  def clear_socket_buffer(gripper_socket="1", read_timeout = 0.1):
      rq_comm_clear_socket_buffer_enabled[rq_socket_to_index(gripper_socket)] = True
  end

  def rq_gripper_id_to_ascii(gripper_id):
      if(gripper_id == "1"):
          return 57
      elif(gripper_id == "2"):
          return 50
      elif(gripper_id == "3"):
          return 51
      elif(gripper_id == "4"):
          return 52
      end
  end

      def scale(value, rawRange, scaledRange):
          def computeSlope(inputRange, outputRange):
              outputRangeDelta = outputRange[1] - outputRange[0]
              inputRangeDelta = inputRange[1] - inputRange[0]

              if (inputRangeDelta == 0):
                  return 0
              else:
                  return outputRangeDelta / inputRangeDelta
              end
          end

          def computeIntercept(slope, inputRange, outputRange):
              return outputRange[0] - (slope * inputRange[0])
          end

          def clipScaledValue(outputScaledValue, outputRange):
              if (outputRange[0] < outputRange[1]):
                  return clipWhenLowerLimitIsLessThanHigher(outputScaledValue, outputRange)
              else:
                  return clipWhenLowerLimitIsGreaterThanHigherLimit(outputScaledValue, outputRange)
              end
          end

          def clipWhenLowerLimitIsGreaterThanHigherLimit(outputScaledValue, outputRange):
              if (outputScaledValue < outputRange[1]):
                  return outputRange[1]
              elif (outputScaledValue > outputRange[0]):
                  return outputRange[0]
              else:
                  return outputScaledValue
              end
          end

          def clipWhenLowerLimitIsLessThanHigher(outputScaledValue, outputRange):
              if (outputScaledValue < outputRange[0]):
                  return outputRange[0]
              elif (outputScaledValue > outputRange[1]):
                  return outputRange[1]
              else:
                  return outputScaledValue
              end
          end

          slope = computeSlope(rawRange, scaledRange)
          intercept = computeIntercept(slope, rawRange, scaledRange)
          scaledValue = slope * value + intercept
          return clipScaledValue(scaledValue, scaledRange)
      end

      def limit(value, range):
          return scale(value, range, range)
      end


  rq_init_comm_if_connected(9, "1")
  rq_init_comm_if_connected(2, "2")
  rq_init_comm_if_connected(3, "3")
  rq_init_comm_if_connected(4, "4")
  rq_print_connected_grippers()
  rq_gripper_communication_thread = run rq_gripper_communication()
  set_closed_norm(97.6470588235294, "1")
  set_open_norm(1.1764705882352942, "1")
  set_closed_mm(0.0, "1")
  set_open_mm(53.0, "1")
  set_closed_norm(100.0, "2")
  set_open_norm(0.0, "2")
  set_closed_mm(0.0, "2")
  set_open_mm(50.0, "2")
  set_closed_norm(100.0, "3")
  set_open_norm(0.0, "3")
  set_closed_mm(0.0, "3")
  set_open_mm(50.0, "3")
  set_closed_norm(100.0, "4")
  set_open_norm(0.0, "4")
  set_closed_mm(0.0, "4")
  set_open_mm(50.0, "4")
  rq_current_limit_enabled = False
  while(not rq_gripper_communication_thread_started):
      sleep(0.008)
  end
  # end: URCap Installation Node
  global AMR_Position=struct(position_identifier=0, x1=0, x2=0, y1=0, y2=0, theta1=0, theta2=0)
  global CAM_Pose=p[0,0,0,0,0,0]
  global CAM_Relation=""
  global CMD_Abort=  False
  global CMD_Clear=  False
  global CMD_Reset=  False
  global CMD_Start=  False
  global CMD_Suspend=  False
  global CMD_Unhold=  False
  global CMD_Unsuspend=  False
  global CNT_Rack_Output=0
  global FNC_Freedrive=  False
  global PRC_TubCounter=0
  global STP=0
  global easyPickCount_4=0
  global easyPickCount_7=0
  global easyPickNoObj_4=0
  global easyPickNoObj_7=0
  global easyPickParts_4=0
  global easyPickParts_7=0
  global TMR_Barcode=0
  global Container_mid_1_p=p[-.379239199143, -.127191311915, .299999999998, .000000000046, -.000000000021, -1.247199999994]
  global Container_mid_1_q=[-2.477408934449926, -1.2969853503591224, -1.875639182904262, -1.539621866126728, 1.5731943360401213, -2.8009955944022717]
  global trigger_otw_p=p[-.364831738276, -.163967193938, .343299997821, .000000000046, -.000000000020, -1.148401333327]
  global trigger_otw_q=[-2.378283213085033, -1.2994862387706814, -1.7634300687554951, -1.6493302004167063, 1.573123683454141, -2.8011223671816943]
  global Waypoint_54_p=p[.008800512419, -.547926542621, .402696567415, -.589884378425, -.007228654778, -.061268144704]
  global Waypoint_54_q=[-1.2044575850116175, -1.3416667741588135, -1.8272563219070435, -0.9884541195682068, 1.3621035814285278, -2.7712565104113978]
  global Waypoint_77_p=p[-.178371829612, -.433927395311, .368082383916, -.086593488055, .704679941724, -.007869906074]
  global Waypoint_77_q=[-1.265390698109762, -1.3355963987163086, -1.7944865226745605, -1.7402602634825648, 0.8780410885810852, -2.7713127771960657]
  global Waypoint_83_p=p[.008800512419, -.547926542621, .402696567415, -.589884378425, -.007228654778, -.061268144704]
  global Waypoint_83_q=[-1.2044575850116175, -1.3416667741588135, -1.8272563219070435, -0.9884541195682068, 1.3621035814285278, -2.7712565104113978]
  global Waypoint_84_p=p[-.178371829612, -.433927395311, .368082383916, -.086593488055, .704679941724, -.007869906074]
  global Waypoint_84_q=[-1.265390698109762, -1.3355963987163086, -1.7944865226745605, -1.7402602634825648, 0.8780410885810852, -2.7713127771960657]
  global Vial_above_1_p=p[.017105793010, -.652093028359, .184920586844, .000000000272, .000000000270, 1.564063451276]
  global Vial_above_1_q=[-1.3375440709712851, -1.9618096977868804, -1.4665759083780685, -1.2837941559171444, 1.5732503672317195, -4.47276330421513]
  global Vial_pick_poi_1_p=p[.017105792852, -.648922724010, .093307568731, .000000000271, .000000000270, 1.564063451276]
  global Vial_pick_poi_1_q=[-1.3366329456391917, -2.0375277831965413, -1.6071432798879028, -1.0675084332049813, 1.57309887265915, -4.471135348858068]
  global Waypoint_86_p=p[.019227646885, -.648669633640, .184920586950, .000000000000, .000000000000, .024063451426]
  global Waypoint_86_q=[-1.3331129109407733, -1.9540750545686123, -1.4775914902901128, -1.280581784992414, 1.5733500744865856, -2.928303704452631]
  global Waypoint_87_p=p[-.032361834699, -.348336136197, .391475576335, -.000008499254, .000014589902, -.004651426820]
  global Waypoint_87_q=[-1.2709335019096129, -1.1914598663441005, -1.708995335060501, -1.8117888533498316, 1.5729683532263925, -2.8379347397710237]
  global Vial_3FG_plac_1_p=p[-.031858676359, -.349402499566, .145301120695, .000000000000, .000000000000, .000000000000]
  global Vial_3FG_plac_1_q=[-1.2723975525801707, -1.252376585823825, -2.3128114007049496, -1.1470592278900167, 1.5730548099411423, -2.8414815174610535]
  global Waypoint_88_p=p[-.032361834699, -.348336136197, .391475576335, -.000008499254, .000014589902, -.004651426820]
  global Waypoint_88_q=[-1.2709335019096129, -1.1914598663441005, -1.708995335060501, -1.8117888533498316, 1.5729683532263925, -2.8379347397710237]
  global cap_dump_1_p=p[-.139168676487, -.420163541420, .146096395183, .000000000000, .000000000000, .000000000000]
  global cap_dump_1_q=[-1.584588644510994, -1.5093464179777323, -2.1118449369620347, -1.091059703602438, 1.5728943834877336, -3.154014906686923]
  global Waypoint_89_p=p[-.032361834699, -.348336136197, .391475576335, -.000008499254, .000014589902, -.004651426820]
  global Waypoint_89_q=[-1.2709335019096129, -1.1914598663441005, -1.708995335060501, -1.8117888533498316, 1.5729683532263925, -2.8379347397710237]
  global Vial_3FG_plac_2_p=p[-.031858676359, -.349402499566, .145301120695, .000000000000, .000000000000, .000000000000]
  global Vial_3FG_plac_2_q=[-1.2723975525801707, -1.252376585823825, -2.3128114007049496, -1.1470592278900167, 1.5730548099411423, -2.8414815174610535]
  global Waypoint_90_p=p[-.032361834699, -.348336136197, .391475576335, -.000008499254, .000014589902, -.004651426820]
  global Waypoint_90_q=[-1.2709335019096129, -1.1914598663441005, -1.708995335060501, -1.8117888533498316, 1.5729683532263925, -2.8379347397710237]
  global cap_dump_2_p=p[-.139168676487, -.420163541420, .146096395183, .000000000000, .000000000000, .000000000000]
  global cap_dump_2_q=[-1.584588644510994, -1.5093464179777323, -2.1118449369620347, -1.091059703602438, 1.5728943834877336, -3.154014906686923]
  global Waypoint_91_p=p[-.032361834699, -.348336136197, .391475576335, -.000008499254, .000014589902, -.004651426820]
  global Waypoint_91_q=[-1.2709335019096129, -1.1914598663441005, -1.708995335060501, -1.8117888533498316, 1.5729683532263925, -2.8379347397710237]
  global Vial_liq_abov_1_p=p[-.025303660977, -.338758622354, .426628485936, -1.315858642253, .800043520260, -.928295855026]
  global Vial_liq_abov_1_q=[-0.3789628187762659, -1.5149522957256814, -2.263045310974121, 0.7870649534412841, -0.750984017048971, -3.2237566153155726]
  global Vial_liq_pick_3_p=p[-.002660428945, -.335984893034, .159389832934, -1.150456778400, .673175527684, -1.010612657503]
  global Vial_liq_pick_3_q=[-0.3660772482501429, -1.4503649038127442, -2.4056053161621094, -1.994692941705221, 0.8039668202400208, -0.2508929411517542]
  global Vial_liq_pick_4_p=p[-.041402486291, -.356791603314, .125395323246, -1.143483969075, .651070210027, -.878721885453]
  global Vial_liq_pick_4_q=[-0.4426233705502476, -1.437252121513727, -2.551930962114307, -1.776528229806984, 0.6562026234073748, -0.43018811960029524]
  global Vial_liq_abov_2_p=p[-.025303660977, -.338758622354, .426628485936, -1.315858642253, .800043520260, -.928295855026]
  global Vial_liq_abov_2_q=[-0.3789628187762659, -1.5149522957256814, -2.263045310974121, 0.7870649534412841, -0.750984017048971, -3.2237566153155726]
  global Liquid_midway_1_p=p[.057575295009, -.583081747994, .306414980749, -1.351675548728, .120935756539, -.096908606303]
  global Liquid_midway_1_q=[-0.895174805318014, -1.7035466633238734, -2.380953073501587, 0.631549521083496, 0.7706599235534668, -2.9455552736865442]
  global shake_3_p=p[.057574880217, -.583085370269, .306422893466, -1.360996190983, -.155555042453, -.438136255921]
  global shake_3_q=[-0.8951800505267542, -1.7035466633238734, -2.380937099456787, 0.6315542894550782, 0.7706599235534669, -2.5394540616517496]
  global shake_4_p=p[.057581636113, -.583090570002, .306439684073, -1.308767904323, .368530312677, .214926493520]
  global shake_4_q=[-0.8951714674579065, -1.7035395107665003, -2.380906343460083, 0.6315504747578125, 0.7706480026245118, -3.3161255787892268]
  global drop_above_3_p=p[.268235025993, -.467784390499, .226219872376, -1.027832627524, -.430841408251, 1.004603115937]
  global drop_above_3_q=[-0.935645882283346, -1.6663371525206507, -2.4252893924713135, 0.41966931402172847, 1.8470635414123535, -3.4600217978106897]
  global drop_above_4_p=p[.219042229014, -.470775657081, .133754190740, -.313004595901, -.344395319364, 1.500564994056]
  global drop_above_4_q=[-1.0601594887284795, -1.70046459045642, -2.0799996233759863, -0.7243227230676759, 1.9429634314685202, -4.115129153870795]
  global liq_tran_3_p=p[.213067510942, -.469567035397, .100231043184, .251862243732, .217902579404, 1.592812335393]
  global liq_tran_3_q=[-0.7789645168037476, -1.822364827406652, -1.8643518410805573, -1.252158963840138, 1.3768134449520435, -3.9328333233290254]
  global drop_above_5_p=p[.219042229014, -.470775657081, .133754190740, -.313004595901, -.344395319364, 1.500564994056]
  global drop_above_5_q=[-1.0601594887284795, -1.70046459045642, -2.0799996233759863, -0.7243227230676759, 1.9429634314685202, -4.115129153870795]
  global Waypoint_92_p=p[.187119460405, -.493959476151, .133754190608, -.313004596540, -.344395317757, 1.500564993991]
  global Waypoint_92_q=[-1.1418328121400876, -1.7310553375189475, -2.033634768766424, -0.772026910513711, 1.958578934631971, -4.201588449364511]
  global liq_tran_4_p=p[.195957706507, -.493022614126, .100231042689, .160718757180, .109807038912, 1.525321508623]
  global liq_tran_4_q=[-0.881740380645474, -1.8244526267589851, -1.865100964490387, -1.1608866323693583, 1.4631433601076713, -3.973915130363038]
  global drop_above_6_p=p[.219042229014, -.470775657081, .133754190740, -.313004595901, -.344395319364, 1.500564994056]
  global drop_above_6_q=[-1.0601594887284795, -1.70046459045642, -2.0799996233759863, -0.7243227230676759, 1.9429634314685202, -4.115129153870795]
  global drop_above_7_p=p[.268235025993, -.467784390499, .226219872376, -1.027832627524, -.430841408251, 1.004603115937]
  global drop_above_7_q=[-0.935645882283346, -1.6663371525206507, -2.4252893924713135, 0.41966931402172847, 1.8470635414123535, -3.4600217978106897]
  global Liquid_midway_2_p=p[.057575295009, -.583081747994, .306414980749, -1.351675548728, .120935756539, -.096908606303]
  global Liquid_midway_2_q=[-0.895174805318014, -1.7035466633238734, -2.380953073501587, 0.631549521083496, 0.7706599235534668, -2.9455552736865442]
  global Vial_drop_abo_1_p=p[.000324902251, -.648569523142, .221894115667, -.873462921366, 1.165852672573, -1.482720593185]
  global Vial_drop_abo_1_q=[-1.0576906334721352, -2.393016994184633, -0.9236232851859159, -2.5729213042279273, 0.7903331288549689, -0.33286325848155585]
  global Vial_liq_drop_1_p=p[.001020867953, -.647659915585, .092915870838, -.834762611599, 1.081942994823, -1.540647900176]
  global Vial_liq_drop_1_q=[-1.0631954168193474, -2.4447642951220825, -1.128811017825127, -2.1983115491972294, 0.8130148661460634, -0.38984988696911316]
  global Vial_drop_abo_2_p=p[.000324902251, -.648569523142, .221894115667, -.873462921366, 1.165852672573, -1.482720593185]
  global Vial_drop_abo_2_q=[-1.0576906334721352, -2.393016994184633, -0.9236232851859159, -2.5729213042279273, 0.7903331288549689, -0.33286325848155585]
  global Spatula_otw_p=p[-.038472058237, -.263141484147, .425351216717, -.000441582511, -.000128175490, 3.034387645854]
  global Spatula_otw_q=[-1.1888947506684495, -1.0083288774886814, -1.7052227056065874, -1.9984805067363443, 1.5730180972985317, 0.48793409320312264]
  global pick_spat_L_abv_p=p[.239059466375, -.067212518441, .280720723617, .000017217488, -.000484427718, 3.106837214660]
  global pick_spat_L_abv_q=[0.292765616142962, -0.8565557553273315, -2.140199892763044, -1.715349495646084, 1.573623142106424, 1.8984976776985687]
  global spat_L_pick_p=p[.242468789885, -.067301915011, .193171208067, .000017217488, -.000484427718, 3.106837214657]
  global spat_L_pick_q=[0.2867414378807389, -0.8600077002089179, -2.3629148016312627, -1.4891831672860159, 1.5737695566221115, 1.8933890858591198]
  global spat_L_lift_p=p[.245402002494, -.067432373551, .289049296496, .000017217490, -.000484427724, 3.106837214657]
  global spat_L_lift_q=[0.2834351187564135, -0.8798320076811592, -2.1119436738532986, -1.7203314352121302, 1.573588313403067, 1.8891054681654005]
  global spat_L_side_p=p[.247133573905, -.017633681797, .289062935631, .000017217490, -.000484427724, 3.106837214657]
  global spat_L_side_q=[0.49719173575848863, -0.8582398211168538, -2.1182130454788215, -1.735610316654931, 1.5735817737572706, 2.1028402698705397]
  global spat_L_up_p=p[.247135508752, -.017665230822, .397130746165, .000017217490, -.000484427724, 3.106837214657]
  global spat_L_up_q=[0.49854946074076967, -0.9346239623559676, -1.808280269374471, -1.969158816463132, 1.5731020084036995, 2.1031742024348157]
  global spat_M_up_p=p[.244670000000, -.112000000000, .420343789747, .000026293990, -.000477463070, 3.067686800857]
  global spat_M_up_q=[0.09097498152209688, -1.0114245603211778, -1.718034632879454, -1.9826932847219538, 1.5730130135866505, 1.734554438783734]
  global spat_M_pick_p=p[.244673518506, -.111985070134, .192299022723, .000043885692, -.000001622442, 3.067686841404]
  global spat_M_pick_q=[0.08868170265231701, -0.9271392933223233, -2.343826449241451, -1.441236864368305, 1.5733923850045939, 1.7345552462242537]
  global spat_S_Up_7_p=p[.243228810603, -.161948321982, .423281604617, .000026293955, -.000477463064, 3.067686800854]
  global spat_S_Up_7_q=[-0.11182322368059516, -1.0716267311491734, -1.6854498186860427, -1.955120134033855, 1.5730106579635699, 1.5317349120701778]
  global spat_S_Pick_4_p=p[.245377020686, -.158668022535, .192285730279, .000026293985, -.000477463062, 3.067686800840]
  global spat_S_Pick_4_q=[-0.10087203759495189, -1.011188488703386, -2.311978084495874, -1.3890267520590838, 1.5735990551056096, 1.5450562970948172]
  global spat_S_Up_8_p=p[.252087445596, -.159242094834, .423281604617, .000026293954, -.000477463070, 3.067686800855]
  global spat_S_Up_8_q=[-0.09804692328730358, -1.0862987822056382, -1.6788706463996483, -1.9470242450550348, 1.5730147401359813, 1.5455107082823842]
  global spat_flatM_up_p=p[.241028517126, -.208127630016, .404671074680, .000026293951, -.000477463078, 3.067686800891]
  global spat_flatM_up_q=[-0.27878462628263456, -1.1217510366315881, -1.7121530048618725, -1.8783279876432832, 1.5731053960668042, 1.3649536117980254]
  global spat_flatM_pick_p=p[.241028983327, -.208057297586, .192270533170, .000026293950, -.000477463079, 3.067686800885]
  global spat_flatM_pick_q=[-0.2805687960562633, -1.1003763929487214, -2.271431297337675, -1.3404236887924883, 1.5734924238720627, 1.3653813047742556]
  global spat_flatS_up_p=p[.237651953780, -.253943828614, .403961222825, .000026293950, -.000477463092, 3.067686800841]
  global spat_flatS_up_q=[-0.42363550926974103, -1.1939944599502539, -1.6745915127240307, -1.843675057902054, 1.5731001874678698, 1.220082820532415]
  global spat_flatS_pick_p=p[.241325662334, -.251726327528, .192256842740, .000026293947, -.000477463087, 3.067686800841]
  global spat_flatS_pick_q=[-0.4144907797170738, -1.1967447109013012, -2.21926362252748, -1.2962499335425761, 1.5733885098427622, 1.2314402238866728]
  global spat_S_pick_p=p[.241585614619, -.158882677087, .191636172448, .000019478956, -.000483249177, 3.097147973434]
  global spat_S_pick_q=[-0.10320942227973173, -1.0007485193115802, -2.317947069452162, -1.3934956127505886, 1.5736112980229278, 1.5132597021160705]
  global spat_S_up_p=p[.248189103503, -.159371150053, .417088864416, .000026293966, -.000477463070, 3.067686800840]
  global spat_S_up_q=[-0.10007737460061872, -1.0730270029702904, -1.7018049146034766, -1.9373622285571734, 1.573045444550866, 1.5435422173047084]
  global Waypoint_7_p=p[-.472820924474, .292439826233, .207418370237, -.137787250486, 2.177332259632, -2.152029714756]
  global Waypoint_7_q=[-2.911134078210732, -1.90240864358569, -1.968768330510411, -2.500365101593811, 0.11427687110891149, 0.0958980389250167]
  global Waypoint_8_p=p[-.357612884176, -.251084817998, .212379799667, -.858181193174, 1.714832512191, -1.687547565568]
  global Waypoint_8_q=[-1.620834863369681, -1.8936194567376496, -1.9821394403832038, -2.4599791457905273, 0.6296693672615152, 0.07625365420707819]
  global Decapp_above_3_p=p[-.013480295948, -.359153355979, .266194408367, -.879653555922, 1.646336924805, -1.709111068605]
  global Decapp_above_3_q=[-0.9632157249872035, -2.0163405763031657, -1.5968194594157152, -2.6579215719847085, 1.251243398585566, 0.047906446502667066]
  global Decapp_place_3_p=p[-.013480295890, -.359153356055, .160907502384, -.879653554902, 1.646336919740, -1.709111066456]
  global Decapp_place_3_q=[-0.9633402410919709, -2.1541179572356635, -1.6937729380888573, -2.4232786481058053, 1.2517342187662468, 0.04818402956922263]
  global Decapp_above_4_p=p[-.013480295948, -.359153355979, .266194408367, -.879653555922, 1.646336924805, -1.709111068605]
  global Decapp_above_4_q=[-0.9632157249872035, -2.0163405763031657, -1.5968194594157152, -2.6579215719847085, 1.251243398585566, 0.047906446502667066]
  global Waypoint_78_p=p[-.051450028091, -.519555688329, .365718563414, -1.287302938145, 1.077637394477, -1.218524965834]
  global Waypoint_78_q=[-0.9214276262416012, -1.8899696965062578, -1.4939326452510562, -2.840015661555725, 0.5585157189668353, 0.033997638875617575]
  global Waypoint_10_p=p[-.466751210260, .252836712095, .259921246286, 1.042686976164, .439333316918, -1.691967798809]
  global Waypoint_10_q=[-3.022216346250036, -1.8383597675135919, -1.566977059184386, -2.046864464116096, 0.8487467526238, -2.4392912369481916]
  global Waypoint_9_p=p[-.538777454962, .370695704977, .175030018143, -.317104215445, 2.082346543003, -2.037631421082]
  global Waypoint_9_q=[-3.1158871966457857, -1.998548595120492, -1.941797010061462, -2.2703530575838844, -0.27573365931009164, -0.06926782177267654]
  global Powder_wayp1_p=p[-.472820924474, .292439826233, .207418370237, -.137787250486, 2.177332259632, -2.152029714756]
  global Powder_wayp1_q=[-2.911134078210732, -1.90240864358569, -1.968768330510411, -2.500365101593811, 0.11427687110891149, 0.0958980389250167]
  global Waypoint_2_p=p[-.357612884176, -.251084817998, .212379799667, -.858181193174, 1.714832512191, -1.687547565568]
  global Waypoint_2_q=[-1.620834863369681, -1.8936194567376496, -1.9821394403832038, -2.4599791457905273, 0.6296693672615152, 0.07625365420707819]
  global Postions_otw_p=p[-.010896578244, -.533368729951, .288851175116, -1.233738470894, 1.195331112012, -1.207314088469]
  global Postions_otw_q=[-0.898791023514228, -2.078490033037677, -1.4499891355755317, -2.7624416226992476, 0.6570218891920963, 0.02136606178275929]
  global cont_A_otw_p=p[.070238108556, -.655257851554, .184611566008, -1.090601381517, 1.404822685081, -1.413645380264]
  global cont_A_otw_q=[-0.990969136335913, -2.7123780097559784, -0.5772671651193146, -3.0005537851220403, 0.84719335943793, 0.020652463706785973]
  global cont_B_otw_p=p[.255895686750, -.501120003087, .157855243207, -1.209177187561, 1.209243088037, -1.209202949417]
  global cont_B_otw_q=[-0.5819602570351563, -2.5181180937953833, -1.0264696604583161, -2.7360726814058687, 0.9880932038785559, -0.004134033524621827]
  global cont_B_safe_p=p[.242897168204, -.501733713795, .237745474779, -1.209212324107, 1.209144328638, -1.209309913894]
  global cont_B_safe_q=[-0.5929699566143585, -2.4210115429142114, -0.9949203644592259, -2.8646436479104267, 0.976678899749076, -0.004020526358775811]
  global cont_C_otw_p=p[.319495487998, -.362719410364, .163846736977, -1.233784872294, 1.195277203291, -1.207325031551]
  global cont_C_otw_q=[-0.3611889651645974, -2.404603865546651, -1.2341573845076566, -2.650535279811077, 1.1944844573128257, 0.01638086594640864]
  global Waypoint_1_p=p[-.352029261722, -.424157832422, .472326578019, -.000004407962, .000020663369, -1.529709227737]
  global Waypoint_1_q=[-2.017015745614491, -1.7423968528991196, -1.0053357238485425, -1.9644715035904907, 1.5727249689896, -2.060727852912713]
  global Waypoint_5_p=p[.219993437017, -.447144142811, .462350040687, .000006087494, .000031090075, .000022232405]
  global Waypoint_5_q=[-0.8406239476037944, -1.5982534362206806, -1.1934200873248484, -1.9205794898315975, 1.5727336676986443, -2.4135960466995314]
  global place_2_home_p=p[-.352029261717, -.424157832411, .329197314759, -.000004407962, .000020663369, -1.529709227737]
  global place_2_home_q=[-2.017880982348384, -1.6708952803108668, -1.462293789471877, -1.5790150659586653, 1.5732060241635952, -2.059940179665328]
  global Waypoint_12_p=p[-.812560029877, -.415067232840, .258518340146, -1.257569567036, 1.159670338548, -1.145019586130]
  global Waypoint_12_q=[-2.3224548809497123, -2.3211405271930765, -1.1304722687551445, -2.8155296475017018, -0.8321758827962036, -0.007205995478960503]
  global Waypoint_18_p=p[-.813643087636, -.416224939441, .099970000000, -1.257570310935, 1.159676546330, -1.145010619029]
  global Waypoint_18_q=[-2.322494764677227, -2.501268559301314, -1.239250885783676, -2.5265468980680197, -0.831327849164623, -0.00732105677136996]
  global Waypoint_19_p=p[-.812560029269, -.415067232191, .079455005744, -1.257569567033, 1.159670338546, -1.145019586137]
  global Waypoint_19_q=[-2.3224951834453367, -2.5274729453886575, -1.2489176533831348, -2.4906644180980346, -0.8312252662037514, -0.007338111970053518]
  global TMR_Barcode_is_counting=False
  thread Timer_Thread():
    while (True):
      if (TMR_Barcode_is_counting):
        TMR_Barcode = TMR_Barcode + get_steptime()
      end
      sync()
    end
  end
  run Timer_Thread()
  def Sub_Vision_V18():
    $ 887 "Sub_Vision_V18" "noBreak"
    $ 888 "PreSettings"
    $ 889 "CAM_LM_Detected≔ False "
    global CAM_LM_Detected=  False
    $ 890 "CAM_Captures≔0"
    global CAM_Captures=0
    $ 891 "CAM_Pose≔p[0,0,0,0,0,0]"
    global CAM_Pose=p[0,0,0,0,0,0]
    $ 892 "CAM_LM_Refinmnt≔ False "
    global CAM_LM_Refinmnt=  False
    $ 893 "CAM_LM_Refined≔ False "
    global CAM_LM_Refined=  False
    $ 894 "CAM_LM_Deviatn≔p[0,0,0,0,0,0]"
    global CAM_LM_Deviatn=p[0,0,0,0,0,0]
    $ 895 "CAM_LM_ID≔0"
    global CAM_LM_ID=0
    $ 896 "CAM_Done≔ False "
    global CAM_Done=  False
    $ 897 "CAM_CNT_Obj≔0"
    global CAM_CNT_Obj=0
    $ 898 "CAM_Result = []"
    CAM_Result = []
    $ 899 "OBJ_Detected≔ False "
    global OBJ_Detected=  False
    $ 900 "FRM_Reference≔p[0,0,0,0,0,0]"
    global FRM_Reference=p[0,0,0,0,0,0]
    $ 901 "'=========='"
    # '=========='
    $ 902 "Switch Action"
    switch_1 = Action
    $ 903 "Case 13"
    if (13 == switch_1):
    elif (15 == switch_1):
      $ 1021 "Case 15"
    elif (131 == switch_1):
      $ 1067 "Case 131"
      $ 1068 "Read (SensoPart)"
      $ 1069 "Action_Info≔'search for landmark'"
      global Action_Info="search for landmark"
      $ 1070 "CAM_LM≔CAM_LMs[4]"
      global CAM_LM=CAM_LMs[4]
      $ 1071 "CAM_Relation≔CAM_LM.capture_relation"
      global CAM_Relation=CAM_LM.capture_relation
      $ 1072 "go to capture pose"
      $ 1075 "If ITM_ID≟1 and JIG≟7"
      if (ITM_ID == 1  and  JIG == 7):
        $ 1076 "PSE_T≔uLM_Cap_SSRack"
        global PSE_T=uLM_Cap_SSRack
      else:
        $ 1077 "ElseIf ITM_ID≟5 and JIG≟7"
        if (ITM_ID == 5  and  JIG == 7):
          $ 1078 "PSE_T≔FRM_Cap_SSRack"
          global PSE_T=FRM_Cap_SSRack
        else:
          $ 1081 "ElseIf ITM_ID≟1 and JIG≟15"
          if (ITM_ID == 1 and JIG == 15):
            $ 1082 "MoveJ"
            $ 1083 "Container_mid_1" "breakAfter"
            movej(get_inverse_kin(Container_mid_1_p, qnear=Container_mid_1_q), a=1.3962634015954636, v=1.0471975511965976, r=0.05)
            $ 1085 "PSE_T≔FRM_Container_const"
            global PSE_T=p[-0.5003348223692186,0.35061804815168285,0.41579001388808423,-5.092943187272062E-5,1.0145185065363121E-4,-2.764319258713288]
          else:
            $ 1086 "ElseIf ITM_ID≟1 and JIG≟21"
            if (ITM_ID == 1 and JIG == 21):
              $ 1088 "PSE_T≔FRM_PoTS_const"
              global PSE_T=p[-0.5403054403210852,-0.10910773999775857,0.4828,3.058497512721046E-6,2.3454853329357316E-5,-2.208510541952706]
            else:
              $ 1089 "ElseIf ITM_ID≟1 and JIG≟17"
              if (ITM_ID == 1 and JIG == 17):
                $ 1090 "MoveJ"
                $ 1091 "zero_scale()"
                zero_scale()
                $ 1092 "trigger_otw" "breakAfter"
                movej(get_inverse_kin(trigger_otw_p, qnear=trigger_otw_q), a=1.3962634015954636, v=1.0471975511965976, r=0.05)
                $ 1096 "PSE_T≔FRM_weigh_scale_const"
                global PSE_T=p[-0.3804866881697204,0.025744252835212,0.4723487455232425,-1.0445769542396123E-4,-1.924788411074358E-5,-2.1691978730572363]
              end
            end
          end
        end
      end
      $ 1097 "do_transition(PSE_T, keep_rxry=False)"
      do_transition(PSE_T, keep_rxry=False)
      $ 1098 "Set"
      set_tcp(p[0.0,0.0,0.161,3.1415,0.0,0.0])
      $ 1099 "MoveJ"
      $ 1100 "PSE_T" "breakAfter"
      movej(PSE_T, a=1.3962634015954636, v=1.7453292519943295)
      $ 1101 "CAM_Pose≔get_actual_tcp_pose()"
      global CAM_Pose= get_actual_tcp_pose ()
      $ 1102 "Loop  not CAM_Done and  not ERROR.FLAG and  not CMD_Stop"
      while (  not  CAM_Done  and    not  ERROR.FLAG  and    not  CMD_Stop):
        $ 1103 "adjust capture pose"
        $ 1104 "If CAM_LM_Detected and CAM_LM_Refinmnt"
        if (CAM_LM_Detected  and  CAM_LM_Refinmnt):
          $ 1105 "PSE_T≔p[0,0,0.300,0,0,0]"
          global PSE_T=p[0,0,0.300,0,0,0]
          $ 1106 "CAM_Pose≔PSE_T"
          global CAM_Pose=PSE_T
          $ 1107 "If  not is_reachable(FRM_Reference,[PSE_T])"
          if (  not  is_reachable(FRM_Reference,[PSE_T])):
            $ 1108 "Error"
            $ 1109 "set_error(ERROR_POSE_NOT_REACHABLE)"
            set_error(ERROR_POSE_NOT_REACHABLE)
          end
          $ 1110 "If  not ERROR.FLAG"
          if (  not  ERROR.FLAG):
            $ 1111 "MoveJ"
            $ 1112 "PSE_T" "breakAfter"
            set_tcp(p[0.0,0.0,0.161,0.0,0.0,0.0])
            movej(pose_trans(FRM_Reference, PSE_T), a=0.8726646259971648, v=1.3962634015954636)
            $ 1113 "CAM_LM_Refined≔ True "
            global CAM_LM_Refined=  True
          end
        else:
          $ 1114 "ElseIf  not CAM_LM_Detected and CAM_Captures>0"
          if (  not  CAM_LM_Detected  and  CAM_Captures>0):
            $ 1115 "MoveL"
            $ 1116 "If FRM_Reference≟p[0,0,0,0,0,0]"
            if (FRM_Reference == p[0,0,0,0,0,0]):
              $ 1117 "PSE_T≔get_random_pose(pose_ref=CAM_Pose, mode='cubic', range_max=[0.150,0.150,0.015])"
              global PSE_T=get_random_pose(pose_ref=CAM_Pose, mode="cubic", range_max=[0.150,0.150,0.015])
            else:
              $ 1122 "Else" "noBreak"
              $ 1123 "PSE_T≔get_random_pose(pose_ref=CAM_Pose, mode='rotation', range_max=[10,10,0])"
              global PSE_T=get_random_pose(pose_ref=CAM_Pose, mode="rotation", range_max=[10,10,0])
              $ 1124 "CAM_LM_Refined≔ True "
              global CAM_LM_Refined=  True
            end
            $ 1125 "If get_inverse_kin_has_solution(pose_trans(FRM_Reference, PSE_T))"
            if (get_inverse_kin_has_solution( pose_trans (FRM_Reference, PSE_T))):
              $ 1126 "Comment"
              # Comment
              $ 1127 "PSE_T" "breakAfter"
              set_tcp(p[0.0,0.0,0.161,3.1415,0.0,0.0])
              movel(pose_trans(FRM_Reference, PSE_T), a=0.03, v=0.05)
            else:
              $ 1128 "Else" "noBreak"
              $ 1129 "'If random pose is out of reach, set the initial cam pose'"
              # 'If random pose is out of reach, set the initial cam pose'
              $ 1130 "PSE_T≔CAM_Pose"
              global PSE_T=CAM_Pose
            end
          end
        end
        $ 1131 "Wait: 2.0"
        sleep(2.0)
        $ 1132 "trigger"
        $ 1133 "If ITM_ID≟1 and JIG≟7"
        if (ITM_ID == 1  and  JIG == 7):
          # begin: URCap Program Node
          #   Source: SensoPart VISOR Robotic, 2.0.6, SensoPart Industriesensorik GmbH
          #   Type: VISOR Trigger
          $ 1134 "# 1 VISOR Trigger"
          visor_changeJob(1, "Landmark_INVITE_2", 6000)
          visor_trigger(1, 6000, "arm")
          # end: URCap Program Node
        else:
          $ 1135 "ElseIf ITM_ID≟5 and JIG≟7"
          if (ITM_ID == 5  and  JIG == 7):
            # begin: URCap Program Node
            #   Source: SensoPart VISOR Robotic, 2.0.6, SensoPart Industriesensorik GmbH
            #   Type: VISOR Trigger
            $ 1136 "# 1 VISOR Trigger"
            visor_changeJob(1, "Landmark_INVITE_2", 6000)
            visor_trigger(1, 6000, "arm")
            # end: URCap Program Node
          else:
            $ 1137 "ElseIf ITM_ID≟13 and JIG≟7"
            if (ITM_ID == 13  and  JIG == 7):
              # begin: URCap Program Node
              #   Source: SensoPart VISOR Robotic, 2.0.6, SensoPart Industriesensorik GmbH
              #   Type: VISOR Trigger
              $ 1138 "# 1 VISOR Trigger"
              visor_changeJob(1, "Landmark_INVITE_2", 6000)
              visor_trigger(1, 6000, "arm")
              # end: URCap Program Node
            else:
              $ 1139 "ElseIf ITM_ID≟1 and JIG≟15"
              if (ITM_ID == 1 and JIG == 15):
                # begin: URCap Program Node
                #   Source: SensoPart VISOR Robotic, 2.0.6, SensoPart Industriesensorik GmbH
                #   Type: VISOR Trigger
                $ 1140 "# 1 VISOR Trigger"
                visor_changeJob(1, "Aztec_no_dot_pick", 6000)
                visor_trigger(1, 6000, "arm")
                # end: URCap Program Node
              else:
                $ 1141 "ElseIf ITM_ID≟1 and JIG≟21"
                if (ITM_ID == 1 and JIG == 21):
                  # begin: URCap Program Node
                  #   Source: SensoPart VISOR Robotic, 2.0.6, SensoPart Industriesensorik GmbH
                  #   Type: VISOR Trigger
                  $ 1142 "# 1 VISOR Trigger"
                  visor_changeJob(1, "PoTS", 6000)
                  visor_trigger(1, 6000, "arm")
                  # end: URCap Program Node
                else:
                  $ 1143 "ElseIf ITM_ID≟1 and JIG≟17"
                  if (ITM_ID == 1 and JIG == 17):
                    # begin: URCap Program Node
                    #   Source: SensoPart VISOR Robotic, 2.0.6, SensoPart Industriesensorik GmbH
                    #   Type: VISOR Trigger
                    $ 1144 "# 1 VISOR Trigger"
                    visor_changeJob(1, "Weigh_target", 6000)
                    visor_trigger(1, 6000, "arm")
                    # end: URCap Program Node
                  end
                end
              end
            end
          end
        end
        $ 1148 "TM_3D_Found≔visor_partsFound(1)"
        global TM_3D_Found= visor_partsFound (1)
        $ 1150 "If TM_3D_Found>0"
        if (TM_3D_Found>0):
          $ 1151 "CAM_LM_Detected≔ True "
          global CAM_LM_Detected=  True
          $ 1152 "CAM_Captures≔0"
          global CAM_Captures=0
        else:
          $ 1153 "Else" "noBreak"
          $ 1154 "CAM_LM_Detected≔ False "
          global CAM_LM_Detected=  False
          $ 1155 "CAM_Captures≔CAM_Captures+1"
          global CAM_Captures=CAM_Captures+1
        end
        $ 1160 "result"
        $ 1161 "If CAM_LM_Detected"
        if (CAM_LM_Detected):
          $ 1162 "If (CAM_LM_Refinmnt and CAM_LM_Refined) or  not CAM_LM_Refinmnt"
          if ((CAM_LM_Refinmnt  and  CAM_LM_Refined)  or    not  CAM_LM_Refinmnt):
            $ 1220 "If ITM_ID≟1 and JIG≟7"
            if (ITM_ID == 1  and  JIG == 7):
              $ 1221 "CAM_LM_SSRack≔visor_getPose3d(1, 0)"
              global CAM_LM_SSRack= visor_getPose3d (1, 0)
            else:
              $ 1222 "ElseIf ITM_ID≟5 and JIG≟7"
              if (ITM_ID == 5  and  JIG == 7):
                $ 1223 "CAM_LM_SSRack≔visor_getPose3d(1, 0)"
                global CAM_LM_SSRack= visor_getPose3d (1, 0)
              else:
                $ 1226 "ElseIf ITM_ID≟1 and JIG≟15"
                if (ITM_ID == 1 and JIG == 15):
                  $ 1227 "CAM_LM_cont≔visor_getPose3d(1, 0)"
                  global CAM_LM_cont= visor_getPose3d (1, 0)
                  $ 1228 "Trigger≔get_actual_tcp_pose()"
                  global Trigger= get_actual_tcp_pose ()
                else:
                  $ 1229 "ElseIf ITM_ID≟1 and JIG≟21"
                  if (ITM_ID == 1 and JIG == 21):
                    $ 1230 "CAM_LM_cont≔visor_getPose3d(1, 0)"
                    global CAM_LM_cont= visor_getPose3d (1, 0)
                    $ 1231 "Trigger≔get_actual_tcp_pose()"
                    global Trigger= get_actual_tcp_pose ()
                  else:
                    $ 1232 "ElseIf ITM_ID≟1 and JIG≟17"
                    if (ITM_ID == 1 and JIG == 17):
                      $ 1233 "CAM_LM_cont≔visor_getPose3d(1, 0)"
                      global CAM_LM_cont= visor_getPose3d (1, 0)
                      $ 1234 "Trigger≔get_actual_tcp_pose()"
                      global Trigger= get_actual_tcp_pose ()
                    end
                  end
                end
              end
            end
            $ 1235 "CAM_Done≔ True "
            global CAM_Done=  True
          end
        else:
          $ 1236 "ElseIf  not CAM_LM_Detected and CAM_Captures<CAM_PRM_Retries"
          if (  not  CAM_LM_Detected  and  CAM_Captures<CAM_PRM_Retries):
            $ 1237 "CAM_LM_Refined≔ False "
            global CAM_LM_Refined=  False
          else:
            $ 1238 "ElseIf CAM_Captures≥CAM_PRM_Retries"
            if (CAM_Captures >= CAM_PRM_Retries):
              $ 1239 "CAM_Done≔ True "
              global CAM_Done=  True
              $ 1240 "Error"
              $ 1241 "set_error(ERROR_NO_LANDMARK)"
              set_error(ERROR_NO_LANDMARK)
            end
          end
        end
      end
    elif (151 == switch_1):
      $ 1242 "Case 151"
      $ 1243 "Detect (SensoPart)"
      $ 1244 "go to capture pose"
      $ 1245 "FRM_Reference≔FRM_Cap_SSRack"
      global FRM_Reference=FRM_Cap_SSRack
      $ 1246 "PSE_T≔p[0,0,-0.00,0,0,0]"
      global PSE_T=p[0,0,-0.00,0,0,0]
      $ 1247 "do_transition(pose_trans(FRM_Reference, PSE_T), keep_rxry=False)"
      do_transition( pose_trans (FRM_Reference, PSE_T), keep_rxry=False)
      $ 1248 "JNT_Q≔get_actual_joint_positions()"
      global JNT_Q= get_actual_joint_positions ()
      $ 1249 "JNT_Q≔[JNT_Q[0], JNT_Q[1], JNT_Q[2], JNT_Q[3], JNT_Q[4], 0]"
      global JNT_Q=[JNT_Q[0], JNT_Q[1], JNT_Q[2], JNT_Q[3], JNT_Q[4], 0]
      $ 1250 "Set"
      set_tcp(p[0.0,0.0,0.161,3.1415,0.0,0.0])
      $ 1251 "movej(get_inverse_kin(pose_trans(FRM_Reference, PSE_T), qnear=JNT_Q))"
      movej(get_inverse_kin( pose_trans (FRM_Reference, PSE_T), qnear=JNT_Q))
      $ 1252 "CAM_Pose≔pose_trans(pose_inv(FRM_Reference), get_actual_tcp_pose())"
      global CAM_Pose= pose_trans ( pose_inv (FRM_Reference),  get_actual_tcp_pose ())
      $ 1253 "Loop  not CAM_Done and  not ERROR.FLAG and  not CMD_Stop"
      while (  not  CAM_Done  and    not  ERROR.FLAG  and    not  CMD_Stop):
        $ 1254 "If  not OBJ_Detected and CAM_Captures>0"
        if (  not  OBJ_Detected  and  CAM_Captures>0):
          $ 1255 "MoveL"
          $ 1256 "If FRM_Reference≟p[0,0,0,0,0,0]"
          if (FRM_Reference == p[0,0,0,0,0,0]):
            $ 1258 "PSE_T≔get_random_pose(pose_ref=CAM_Pose, mode='rotation', range_max=[15,15,0])"
            global PSE_T=get_random_pose(pose_ref=CAM_Pose, mode="rotation", range_max=[15,15,0])
          else:
            $ 1259 "Else" "noBreak"
            $ 1260 "PSE_T≔get_random_pose(pose_ref=CAM_Pose, mode='rotation', range_max=[10,10,0])"
            global PSE_T=get_random_pose(pose_ref=CAM_Pose, mode="rotation", range_max=[10,10,0])
          end
          $ 1261 "If get_inverse_kin_has_solution(pose_trans(FRM_Reference, PSE_T))"
          if (get_inverse_kin_has_solution( pose_trans (FRM_Reference, PSE_T))):
            $ 1262 "PSE_T" "breakAfter"
            set_tcp(p[0.0,0.0,0.161,3.1415,0.0,0.0])
            movel(pose_trans(FRM_Reference, PSE_T), a=0.03, v=0.05)
          else:
            $ 1263 "Else" "noBreak"
            $ 1264 "'If random pose is out of reach, set the initial cam pose'"
            # 'If random pose is out of reach, set the initial cam pose'
            $ 1265 "PSE_T≔CAM_Pose"
            global PSE_T=CAM_Pose
            $ 1266 "PSE_T" "breakAfter"
            set_tcp(p[0.0,0.0,0.161,3.1415,0.0,0.0])
            movel(pose_trans(FRM_Reference, PSE_T), a=0.03, v=0.05)
          end
        end
        $ 1267 "Wait: 0.5"
        sleep(0.5)
        $ 1268 "Set"
        set_tcp(p[0.0,0.0,0.161,3.1415,0.0,0.0])
        # begin: URCap Program Node
        #   Source: SensoPart VISOR Robotic, 2.0.6, SensoPart Industriesensorik GmbH
        #   Type: VISOR Trigger
        $ 1269 "# 1 VISOR Trigger"
        visor_changeJob(1, "Object Detection Single", 6000)
        visor_trigger(1, 6000, "arm")
        # end: URCap Program Node
        $ 1270 "If visor_isResponseOk(1)"
        if ( visor_isResponseOk (1)):
          $ 1271 "CAM_CNT_Obj≔visor_partsFound(1)"
          global CAM_CNT_Obj= visor_partsFound (1)
          $ 1272 "CAM_OBJ_Pose≔visor_getPose3d(1, 0)"
          global CAM_OBJ_Pose= visor_getPose3d (1, 0)
          $ 1273 "If CAM_CNT_Obj>0"
          if (CAM_CNT_Obj>0):
            $ 1274 "CAM_OBJ_Color≔visor_getAdditionalData(1, 0)"
            global CAM_OBJ_Color= visor_getAdditionalData (1, 0)
            $ 1275 "CAM_DetectScore≔to_num(visor_getAdditionalData(1, 1))/1000"
            global CAM_DetectScore=to_num( visor_getAdditionalData (1, 1))/1000
            $ 1276 "OBJ_Detected≔ True "
            global OBJ_Detected=  True
          end
        else:
          $ 1277 "Else" "noBreak"
          $ 1278 "CAM_Captures≔CAM_Captures+1"
          global CAM_Captures=CAM_Captures+1
        end
        $ 1279 "If OBJ_Detected"
        if (OBJ_Detected):
          $ 1280 "Get object data"
          $ 1281 "PRC_CntDetect≔0"
          global PRC_CntDetect=0
          $ 1282 "Loop PRC_CntDetect<CAM_CNT_Obj"
          while (PRC_CntDetect<CAM_CNT_Obj):
            $ 1283 "get object and jig number"
            $ 1284 "If ITM_ID≟1 and JIG≟7"
            if (ITM_ID == 1  and  JIG == 7):
              $ 1285 "FRM_Reference≔FRM_Cap_SSRack"
              global FRM_Reference=FRM_Cap_SSRack
            else:
              $ 1286 "ElseIf ITM_ID≟5 and JIG≟7"
              if (ITM_ID == 5  and  JIG == 7):
                $ 1287 "FRM_Reference≔uLM_Cap_SSRack"
                global FRM_Reference=uLM_Cap_SSRack
              end
            end
            $ 1290 "PSE_T≔pose_trans(pose_inv(FRM_Reference), CAM_OBJ_Pose)"
            global PSE_T= pose_trans ( pose_inv (FRM_Reference), CAM_OBJ_Pose)
            $ 1291 "CAM_Result.append(get_pattern_counter(PSE_T, 'X', pattern=[10, 5], patternsize=[0.181, 0.081]))"
            CAM_Result.append(get_pattern_counter(PSE_T, "X", pattern=[10, 5], patternsize=[0.181, 0.081]))
            $ 1292 "PRC_CntDetect≔PRC_CntDetect+1"
            global PRC_CntDetect=PRC_CntDetect+1
          end
          $ 1293 "CAM_Done≔ True "
          global CAM_Done=  True
        else:
          $ 1294 "ElseIf CAM_Captures≥CAM_PRM_Retries"
          if (CAM_Captures >= CAM_PRM_Retries):
            $ 1295 "CAM_Done≔ True "
            global CAM_Done=  True
          else:
            $ 1296 "Else" "noBreak"
            $ 1297 "CAM_Captures≔CAM_Captures+1"
            global CAM_Captures=CAM_Captures+1
          end
        end
      end
    end
    $ 1298 "'=========='"
    # '=========='
    $ 1299 "PostSettings"
    $ 1300 "FRM_Reference≔p[0,0,0,0,0,0]"
    global FRM_Reference=p[0,0,0,0,0,0]
    $ 1301 "Set"
    set_tcp(p[0.0,0.0,0.161,3.1415,0.0,0.0])
    $ 1302 "CAM_Pose≔p[0,0,0,0,0,0]"
    global CAM_Pose=p[0,0,0,0,0,0]
    $ 1303 "Action≔0"
    global Action=0
    $ 1304 "Action_Info≔''"
    global Action_Info=""
  end
  def Sub_AMR_MiR_V3():
    $ 1305 "Sub_AMR_MiR_V3" "noBreak"
    $ 1306 "PreSettings"
    $ 1307 "AMR_TargetList≔[1,2,3,4,5,6,21,22,23,24,31,32,33,34,35,36,37,38,41]"
    global AMR_TargetList=[1,2,3,4,5,6,21,22,23,24,31,32,33,34,35,36,37,38,41]
    $ 1308 "AMR_Done≔ False "
    global AMR_Done=  False
    $ 1309 "AMR_PosActual≔T2O_Current_Pos"
    global AMR_PosActual=modbus_get_signal_status("T2O_Current_Pos")
    $ 1310 "AMR_Attemps≔T2O_Nav_Attemps"
    global AMR_Attemps=modbus_get_signal_status("T2O_Nav_Attemps")
    $ 1311 "AMR_Battery≔MiR_Battery_Lvl"
    global AMR_Battery=modbus_get_signal_status("MiR_Battery_Lvl")
    $ 1312 "AMR_Charging≔(T2O_Charging≟1)"
    global AMR_Charging=(modbus_get_signal_status("T2O_Charging") == 1)
    $ 1313 "AMR_Position≔struct(position_identifier=T2O_Current_Pos, x1=MiR_Position_X1, x2=MiR_Position_X2, y1=MiR_Position_Y1, y2=MiR_Position_Y2, theta1=MiR_Theta_1, theta2=MiR_Theta_2) "
    global AMR_Position=struct(position_identifier=modbus_get_signal_status("T2O_Current_Pos"), x1=modbus_get_signal_status("MiR_Position_X1"), x2=modbus_get_signal_status("MiR_Position_X2"), y1=modbus_get_signal_status("MiR_Position_Y1"), y2=modbus_get_signal_status("MiR_Position_Y2"), theta1=modbus_get_signal_status("MiR_Theta_1"), theta2=modbus_get_signal_status("MiR_Theta_2"))
    $ 1314 "If MiR_Mode≠7"
    if (modbus_get_signal_status("MiR_Mode") != 7):
      $ 1315 "Error"
      $ 1316 "set_error(ERROR_AMR_WRONG_MODE)"
      set_error(ERROR_AMR_WRONG_MODE)
      $ 1317 "AMR_Done≔ True "
      global AMR_Done=  True
    end
    $ 1318 "'=========='"
    # '=========='
    $ 1319 "Switch STATE"
    switch_1 = STATE
    $ 1320 "Case 1"
    if (1 == switch_1):
      $ 1321 "stopping"
      $ 1322 "If T2O_Done≟1 and O2T_Acknowledge≟0"
      if (modbus_get_signal_status("T2O_Done") == 1  and  modbus_get_signal_status("O2T_Acknowledge") == 0):
        $ 1323 "Set O2T_Acknowledge=1"
        modbus_set_output_register("O2T_Acknowledge", 1)
      end
      $ 1324 "Set MiR_CMD_Stop=On"
      modbus_set_output_signal("MiR_CMD_Stop", True)
      $ 1325 "AMR_Position.position_identifier = 0"
      AMR_Position.position_identifier = 0
      $ 1326 "AMR_Done≔ True "
      global AMR_Done=  True
    elif (2 == switch_1):
      $ 1327 "Case 2"
      $ 1328 "stopped"
      $ 1329 "If MiR_State≠3 and MiR_State≠5"
      if (modbus_get_signal_status("MiR_State") != 3  and  modbus_get_signal_status("MiR_State") != 5):
        $ 1330 "Set MiR_CMD_Stop=Off"
        modbus_set_output_signal("MiR_CMD_Stop", False)
      end
    elif (3 == switch_1):
      $ 1331 "Case 3"
      $ 1332 "resetting"
      $ 1333 "Set O2T_Mis_Main=Off"
      modbus_set_output_signal("O2T_Mis_Main", False)
      $ 1334 "Set O2T_Mis_Charge=Off"
      modbus_set_output_signal("O2T_Mis_Charge", False)
      $ 1335 "If MiR_Mis_Queue>0"
      if (modbus_get_signal_status("MiR_Mis_Queue")>0):
        $ 1336 "Set MiR_CMD_Clear_Q=On"
        modbus_set_output_signal("MiR_CMD_Clear_Q", True)
        $ 1337 "Wait MiR_Mis_Queue≟0"
        while (not(modbus_get_signal_status("MiR_Mis_Queue") == 0)):
          sync()
        end
        $ 1338 "Set MiR_CMD_Clear_Q=Off"
        modbus_set_output_signal("MiR_CMD_Clear_Q", False)
      end
      $ 1339 "If MiR_Error_ID≠0"
      if (modbus_get_signal_status("MiR_Error_ID") != 0):
        $ 1340 "Set MiR_CMD_Clear_E=On"
        modbus_set_output_signal("MiR_CMD_Clear_E", True)
        $ 1341 "Wait MiR_Error_ID≟0"
        while (not(modbus_get_signal_status("MiR_Error_ID") == 0)):
          sync()
        end
        $ 1342 "Set MiR_CMD_Clear_E=Off"
        modbus_set_output_signal("MiR_CMD_Clear_E", False)
      end
      $ 1343 "Set O2T_Action=0"
      modbus_set_output_register("O2T_Action", 0)
      $ 1344 "Set O2T_Acknowledge=0"
      modbus_set_output_register("O2T_Acknowledge", 0)
      $ 1345 "Set O2T_Target_Pos=0"
      modbus_set_output_register("O2T_Target_Pos", 0)
      $ 1346 "Set O2T_Footprint=0"
      modbus_set_output_register("O2T_Footprint", 0)
      $ 1347 "Set O2T_ProtectOff=0"
      modbus_set_output_register("O2T_ProtectOff", 0)
      $ 1348 "Set O2T_Dock=0"
      modbus_set_output_register("O2T_Dock", 0)
      $ 1349 "AMR_Attemps≔0"
      global AMR_Attemps=0
      $ 1350 "AMR_PosTarget≔0"
      global AMR_PosTarget=0
      $ 1351 "AMR_Step≔0"
      global AMR_Step=0
      $ 1352 "AMR_AtTarget≔ False "
      global AMR_AtTarget=  False
      $ 1353 "If MiR_State≟4 or MiR_State≟3 or MiR_State≟10"
      if (modbus_get_signal_status("MiR_State") == 4  or  modbus_get_signal_status("MiR_State") == 3  or  modbus_get_signal_status("MiR_State") == 10):
        $ 1354 "AMR_Done≔ True "
        global AMR_Done=  True
      end
    elif (5 == switch_1):
      $ 1355 "Case 5"
      $ 1356 "starting"
      $ 1357 "If MiR_State≟4"
      if (modbus_get_signal_status("MiR_State") == 4):
        $ 1358 "Set MiR_CMD_Start=On"
        modbus_set_output_signal("MiR_CMD_Start", True)
        $ 1359 "Wait MiR_State≠4"
        while (not(modbus_get_signal_status("MiR_State") != 4)):
          sync()
        end
        $ 1360 "Set MiR_CMD_Start=Off"
        modbus_set_output_signal("MiR_CMD_Start", False)
        $ 1361 "AMR_Done≔ True "
        global AMR_Done=  True
      else:
        $ 1362 "ElseIf MiR_State≟10"
        if (modbus_get_signal_status("MiR_State") == 10):
          $ 1363 "'MiR in protective stop. Wait'"
          # 'MiR in protective stop. Wait'
          $ 1364 "AMR_Done≔ True "
          global AMR_Done=  True
        else:
          $ 1365 "ElseIf MiR_State≟3"
          if (modbus_get_signal_status("MiR_State") == 3):
            $ 1366 "AMR_Done≔ True "
            global AMR_Done=  True
          end
        end
      end
    elif (6 == switch_1):
      $ 1367 "Case 6"
      $ 1368 "execute"
      $ 1369 "AMR_AtTarget≔(AMR_PosActual≟AMR_PosTarget)"
      global AMR_AtTarget=(AMR_PosActual == AMR_PosTarget)
      $ 1370 "Switch AMR_Step"
      switch_2 = AMR_Step
      $ 1371 "Case 0"
      if (0 == switch_2):
        $ 1372 "If  not AMR_AtTarget"
        if (  not  AMR_AtTarget):
          $ 1373 "AMR_Step≔1"
          global AMR_Step=1
        else:
          $ 1374 "Else" "noBreak"
          $ 1375 "AMR_Done≔ True "
          global AMR_Done=  True
        end
      elif (1 == switch_2):
        $ 1376 "Case 1"
        $ 1377 "general Settings"
        $ 1378 "Set O2T_Acknowledge=0"
        modbus_set_output_register("O2T_Acknowledge", 0)
        $ 1379 "check for error"
        $ 1380 "If OBJ_Picked and MiR_State≟10"
        if (OBJ_Picked  and  modbus_get_signal_status("MiR_State") == 10):
          $ 1381 "Error"
          $ 1382 "set_error(ERROR_ROBOT_ARM_NOT_IN_HOME_POSE)"
          set_error(ERROR_ROBOT_ARM_NOT_IN_HOME_POSE)
          $ 1383 "Action≔0"
          global Action=0
        else:
          $ 1384 "ElseIf  not found_in_list(AMR_PosTarget, AMR_TargetList)"
          if (  not  found_in_list(AMR_PosTarget, AMR_TargetList)):
            $ 1385 "Error"
            $ 1386 "set_error(ERROR_UNKNOWN_POSE)"
            set_error(ERROR_UNKNOWN_POSE)
            $ 1387 "Action≔0"
            global Action=0
          end
        end
        $ 1388 "If MiR_State≟3"
        if (modbus_get_signal_status("MiR_State") == 3):
          $ 1389 "Set MiR_CMD_Start=Off"
          modbus_set_output_signal("MiR_CMD_Start", False)
          $ 1390 "Switch Action"
          switch_3 = Action
          $ 1391 "Case 51"
          if (51 == switch_3):
            $ 1392 "Charge"
            $ 1393 "'trigger the charging mission'"
            # 'trigger the charging mission'
            $ 1394 "'target pos is predefined'"
            # 'target pos is predefined'
            $ 1395 "Set O2T_Footprint=0"
            modbus_set_output_register("O2T_Footprint", 0)
            $ 1396 "Set O2T_Action=1"
            modbus_set_output_register("O2T_Action", 1)
            $ 1397 "If MiR_Mis_Queue≟0"
            if (modbus_get_signal_status("MiR_Mis_Queue") == 0):
              $ 1398 "Set O2T_Mis_Charge=On"
              modbus_set_output_signal("O2T_Mis_Charge", True)
              $ 1399 "Wait MiR_Mis_Queue≥1"
              while (not(modbus_get_signal_status("MiR_Mis_Queue") >= 1)):
                sync()
              end
              $ 1400 "Set O2T_Mis_Charge=Off"
              modbus_set_output_signal("O2T_Mis_Charge", False)
            end
          elif (52 == switch_3):
            $ 1401 "Case 52"
            $ 1402 "Navigate"
            $ 1403 "'trigger the standard missoin'"
            # 'trigger the standard missoin'
            $ 1404 "Set O2T_Footprint=AMR_FootprintID"
            modbus_set_output_register("O2T_Footprint", AMR_FootprintID)
            $ 1405 "Set O2T_Target_Pos=AMR_PosTarget"
            modbus_set_output_register("O2T_Target_Pos", AMR_PosTarget)
            $ 1406 "Set O2T_Action=2"
            modbus_set_output_register("O2T_Action", 2)
            $ 1407 "If MiR_Mis_Queue≟0"
            if (modbus_get_signal_status("MiR_Mis_Queue") == 0):
              $ 1408 "Set O2T_Mis_Main=On"
              modbus_set_output_signal("O2T_Mis_Main", True)
              $ 1409 "Wait MiR_Mis_Queue≥1"
              while (not(modbus_get_signal_status("MiR_Mis_Queue") >= 1)):
                sync()
              end
              $ 1410 "Set O2T_Mis_Main=Off"
              modbus_set_output_signal("O2T_Mis_Main", False)
            end
          end
        else:
          $ 1411 "ElseIf MiR_State≟4"
          if (modbus_get_signal_status("MiR_State") == 4):
            $ 1412 "Set MiR_CMD_Start=On"
            modbus_set_output_signal("MiR_CMD_Start", True)
          else:
            $ 1413 "ElseIf MiR_State≟5"
            if (modbus_get_signal_status("MiR_State") == 5):
              $ 1414 "AMR_Step≔2"
              global AMR_Step=2
            else:
              $ 1415 "ElseIf MiR_State≟10"
              if (modbus_get_signal_status("MiR_State") == 10):
                $ 1416 "'AMR still in safeguard stop'"
                # 'AMR still in safeguard stop'
              end
            end
          end
        end
      elif (2 == switch_2):
        $ 1417 "Case 2"
        $ 1418 "acknowledge handshake"
        $ 1419 "If T2O_Done≟1 and O2T_Acknowledge≟0"
        if (modbus_get_signal_status("T2O_Done") == 1  and  modbus_get_signal_status("O2T_Acknowledge") == 0):
          $ 1420 "Set O2T_Acknowledge=1"
          modbus_set_output_register("O2T_Acknowledge", 1)
        else:
          $ 1421 "ElseIf T2O_Done≟0 and O2T_Acknowledge≟1"
          if (modbus_get_signal_status("T2O_Done") == 0  and  modbus_get_signal_status("O2T_Acknowledge") == 1):
            $ 1422 "Set O2T_Acknowledge=0"
            modbus_set_output_register("O2T_Acknowledge", 0)
            $ 1423 "AMR_AtTarget≔(AMR_PosActual≟AMR_PosTarget)"
            global AMR_AtTarget=(AMR_PosActual == AMR_PosTarget)
            $ 1424 "AMR_Done≔ True "
            global AMR_Done=  True
          end
        end
      end
      $ 1425 "translate errors"
      $ 1426 "If AMR_Done"
      if (AMR_Done):
        $ 1427 "Switch T2O_Error_ID"
        switch_2 = modbus_get_signal_status("T2O_Error_ID")
        $ 1428 "Case 2003"
        if (2003 == switch_2):
          $ 1429 "error"
          $ 1430 "set_error(ERROR_NOT_DOCKED)"
          set_error(ERROR_NOT_DOCKED)
        elif (2007 == switch_2):
          $ 1431 "Case 2007"
          $ 1432 "error"
          $ 1433 "set_error(ERROR_NOT_REACHABLE_TARGET)"
          set_error(ERROR_NOT_REACHABLE_TARGET)
        elif (2008 == switch_2):
          $ 1434 "Case 2008"
          $ 1435 "error"
          $ 1436 "set_error(ERROR_CHARGING_NOT_STARTED)"
          set_error(ERROR_CHARGING_NOT_STARTED)
        end
      end
    elif (7 == switch_1):
      $ 1437 "Case 7"
      $ 1438 "completing"
      $ 1439 "If MiR_Mis_Queue>0"
      if (modbus_get_signal_status("MiR_Mis_Queue")>0):
        $ 1440 "Set MiR_CMD_Abort=On"
        modbus_set_output_signal("MiR_CMD_Abort", True)
        $ 1441 "Wait MiR_Mis_Queue≟0"
        while (not(modbus_get_signal_status("MiR_Mis_Queue") == 0)):
          sync()
        end
        $ 1442 "Set MiR_CMD_Abort=Off"
        modbus_set_output_signal("MiR_CMD_Abort", False)
      end
      $ 1443 "If MiR_State≟3 or MiR_State≟10"
      if (modbus_get_signal_status("MiR_State") == 3  or  modbus_get_signal_status("MiR_State") == 10):
        $ 1444 "AMR_Done≔ True "
        global AMR_Done=  True
      end
    elif (9 == switch_1):
      $ 1445 "Case 9"
      $ 1446 "holding"
      $ 1447 "Set MiR_CMD_Abort=On"
      modbus_set_output_signal("MiR_CMD_Abort", True)
      $ 1448 "If MiR_State≟3 or MiR_State≟10"
      if (modbus_get_signal_status("MiR_State") == 3  or  modbus_get_signal_status("MiR_State") == 10):
        $ 1449 "Set MiR_CMD_Abort=Off"
        modbus_set_output_signal("MiR_CMD_Abort", False)
        $ 1450 "AMR_Done≔ True "
        global AMR_Done=  True
      end
    elif (11 == switch_1):
      $ 1451 "Case 11"
      $ 1452 "unholding"
      $ 1453 "Set MiR_CMD_Start=On"
      modbus_set_output_signal("MiR_CMD_Start", True)
      $ 1454 "If MiR_State≠4"
      if (modbus_get_signal_status("MiR_State") != 4):
        $ 1455 "Set MiR_CMD_Start=Off"
        modbus_set_output_signal("MiR_CMD_Start", False)
        $ 1456 "AMR_Step≔0"
        global AMR_Step=0
        $ 1457 "AMR_Done≔ True "
        global AMR_Done=  True
      end
    elif (12 == switch_1):
      $ 1458 "Case 12"
      $ 1459 "suspending"
      $ 1460 "'none'"
      # 'none'
    elif (14 == switch_1):
      $ 1461 "Case 14"
      $ 1462 "unsuspending"
      $ 1463 "'none'"
      # 'none'
    elif (15 == switch_1):
      $ 1464 "Case 15"
      $ 1465 "aborting"
      $ 1466 "Set MiR_CMD_Abort=On"
      modbus_set_output_signal("MiR_CMD_Abort", True)
      $ 1467 "Wait MiR_State≟3"
      while (not(modbus_get_signal_status("MiR_State") == 3)):
        sync()
      end
      $ 1468 "Set MiR_CMD_Abort=Off"
      modbus_set_output_signal("MiR_CMD_Abort", False)
    elif (17 == switch_1):
      $ 1469 "Case 17"
      $ 1470 "clearing"
      $ 1471 "If MiR_Error_ID≠0"
      if (modbus_get_signal_status("MiR_Error_ID") != 0):
        $ 1472 "Set MiR_CMD_Clear_E=On"
        modbus_set_output_signal("MiR_CMD_Clear_E", True)
        $ 1473 "Wait MiR_Error_ID≟0"
        while (not(modbus_get_signal_status("MiR_Error_ID") == 0)):
          sync()
        end
        $ 1474 "Set MiR_CMD_Clear_E=Off"
        modbus_set_output_signal("MiR_CMD_Clear_E", False)
      end
      $ 1475 "If MiR_Error_ID≟0"
      if (modbus_get_signal_status("MiR_Error_ID") == 0):
        $ 1476 "AMR_Done≔ True "
        global AMR_Done=  True
      end
    end
    $ 1477 "'=========='"
    # '=========='
    $ 1478 "PostSettings"
    $ 1479 "AMR_Position≔struct(position_identifier=T2O_Current_Pos, x1=MiR_Position_X1, x2=MiR_Position_X2, y1=MiR_Position_Y1, y2=MiR_Position_Y2, theta1=MiR_Theta_1, theta2=MiR_Theta_2) "
    global AMR_Position=struct(position_identifier=modbus_get_signal_status("T2O_Current_Pos"), x1=modbus_get_signal_status("MiR_Position_X1"), x2=modbus_get_signal_status("MiR_Position_X2"), y1=modbus_get_signal_status("MiR_Position_Y1"), y2=modbus_get_signal_status("MiR_Position_Y2"), theta1=modbus_get_signal_status("MiR_Theta_1"), theta2=modbus_get_signal_status("MiR_Theta_2"))
  end
  def Sub_Action_V4():
    $ 1480 "Sub_Action_V4" "noBreak"
    $ 1481 "PreSettings"
    $ 1482 "init poses"
    $ 1483 "PSE_A≔p[0,0,0,0,0,0]"
    global PSE_A=p[0,0,0,0,0,0]
    $ 1484 "PSE_A_H≔p[0,0,0,0,0,0]"
    global PSE_A_H=p[0,0,0,0,0,0]
    $ 1485 "PSE_T≔p[0,0,0,0,0,0]"
    global PSE_T=p[0,0,0,0,0,0]
    $ 1486 "PSE_T_H≔p[0,0,0,0,0,0]"
    global PSE_T_H=p[0,0,0,0,0,0]
    $ 1487 "PSE_G≔p[0,0,0,0,0,0]"
    global PSE_G=p[0,0,0,0,0,0]
    $ 1488 "PSE_G_H≔p[0,0,0,0,0,0]"
    global PSE_G_H=p[0,0,0,0,0,0]
    $ 1489 "PSE_R≔p[0,0,0,0,0,0]"
    global PSE_R=p[0,0,0,0,0,0]
    $ 1490 "PSE_R_H≔p[0,0,0,0,0,0]"
    global PSE_R_H=p[0,0,0,0,0,0]
    $ 1491 "JNT_Q≔[0,0,0,0,0,0]"
    global JNT_Q=[0,0,0,0,0,0]
    $ 1492 "JNT_S≔[0,0,0,0,0,0]"
    global JNT_S=[0,0,0,0,0,0]
    $ 1493 "Gripping parameters"
    $ 1494 "OBJ = find_object_by_type(OBJs, OBJ_Type)"
    OBJ = find_object_by_type(OBJs, OBJ_Type)
    $ 1495 "GRP_Open_Pos≔OBJ.dimension.diameter * 1000 + 6"
    global GRP_Open_Pos=OBJ.dimension.diameter * 1000 + 6
    $ 1496 "GRP_Offset≔OBJ.gripper_offset"
    global GRP_Offset=OBJ.gripper_offset
    $ 1497 "rq_set_force_norm(50)"
     rq_set_force_norm (50)
    $ 1498 "rq_set_speed_norm(50)"
     rq_set_speed_norm (50)
    $ 1499 "Switch ITM_ID"
    switch_1 = ITM_ID
    $ 1500 "Case 1"
    if (1 == switch_1):
      $ 1501 "uML"
      $ 1502 "JIG2 = find_object_by_type(JIGs, JIG)"
      JIG2 = find_object_by_type(JIGs, JIG)
      $ 1503 "JIG_Offset≔JIG2.jig_offset"
      global JIG_Offset=JIG2.jig_offset
      $ 1504 "Switch JIG"
      switch_2 = JIG
      $ 1505 "Case 1"
      if (1 == switch_2):
        $ 1506 "3FG"
        $ 1507 "define poses"
        $ 1508 "FRM_Reference≔ULM_3FG"
        global FRM_Reference=ULM_3FG
        $ 1509 "JNT_Q≔JNT_HOME"
        global JNT_Q=JNT_HOME
        $ 1510 "PSE_T≔pose_trans(GRP_Offset, JIG_Offset)"
        global PSE_T= pose_trans (GRP_Offset, JIG_Offset)
        $ 1511 "PSE_A≔pose_trans(PSE_T, p[0,0,0.100,0,0,0])"
        global PSE_A= pose_trans (PSE_T, p[0,0,0.100,0,0,0])
        $ 1512 "PSE_R≔pose_add(PSE_T, p[0,0,0.100,0,0,0])"
        global PSE_R= pose_add (PSE_T, p[0,0,0.100,0,0,0])
      elif (2 == switch_2):
        $ 1513 "Case 2"
        $ 1514 "Input"
        $ 1515 "'CHANGE THE REFERENCE TO THE FRAME TO MOVE IN'"
        # 'CHANGE THE REFERENCE TO THE FRAME TO MOVE IN'
        $ 1516 "define poses"
        $ 1517 "FRM_Reference≔ULM_Input"
        global FRM_Reference=ULM_Input
        $ 1518 "PSE_T≔pose_trans(pose_trans(get_pattern_pos_rectangle(OBJ_Nbr, 'X', [10,5], patternsize=[0.181,0.081]), GRP_Offset), JIG_Offset)"
        global PSE_T= pose_trans ( pose_trans (get_pattern_pos_rectangle(OBJ_Nbr, "X", [10,5], patternsize=[0.181,0.081]), GRP_Offset), JIG_Offset)
        $ 1519 "If Action≟1"
        if (Action == 1):
          $ 1520 "PSE_R≔pose_add(PSE_T, p[0,0,0.200,0,0,0])"
          global PSE_R= pose_add (PSE_T, p[0,0,0.200,0,0,0])
          $ 1521 "PSE_A≔pose_add(PSE_T, p[0,0,0.100,0,0,0])"
          global PSE_A= pose_add (PSE_T, p[0,0,0.100,0,0,0])
        else:
          $ 1522 "ElseIf Action≟2"
          if (Action == 2):
            $ 1523 "PSE_R≔pose_add(PSE_T, p[0,0,0.100,0,0,0])"
            global PSE_R= pose_add (PSE_T, p[0,0,0.100,0,0,0])
            $ 1524 "PSE_A≔pose_add(PSE_T, p[0,0,0.200,0,0,0])"
            global PSE_A= pose_add (PSE_T, p[0,0,0.200,0,0,0])
          end
        end
      elif (3 == switch_2):
        $ 1525 "Case 3"
        $ 1526 "Output"
        $ 1527 "'CHANGE THE REFERENCE TO THE FRAME TO MOVE IN'"
        # 'CHANGE THE REFERENCE TO THE FRAME TO MOVE IN'
        $ 1528 "define poses"
        $ 1529 "FRM_Reference≔ULM_Output"
        global FRM_Reference=ULM_Output
        $ 1530 "PSE_T≔pose_trans(pose_trans(get_pattern_pos_rectangle(OBJ_Nbr, 'X', [10,5], patternsize=[0.181,0.081]), GRP_Offset), JIG_Offset)"
        global PSE_T= pose_trans ( pose_trans (get_pattern_pos_rectangle(OBJ_Nbr, "X", [10,5], patternsize=[0.181,0.081]), GRP_Offset), JIG_Offset)
        $ 1532 "If Action≟1"
        if (Action == 1):
          $ 1533 "PSE_R≔pose_add(PSE_T, p[0,0,0.200,0,0,0])"
          global PSE_R= pose_add (PSE_T, p[0,0,0.200,0,0,0])
          $ 1534 "PSE_A≔pose_add(PSE_T, p[0,0,0.100,0,0,0])"
          global PSE_A= pose_add (PSE_T, p[0,0,0.100,0,0,0])
        else:
          $ 1535 "ElseIf Action≟2"
          if (Action == 2):
            $ 1536 "PSE_R≔pose_add(PSE_T, p[0,0,0.100,0,0,0])"
            global PSE_R= pose_add (PSE_T, p[0,0,0.100,0,0,0])
            $ 1537 "PSE_A≔pose_add(PSE_T, p[0,0,0.200,0,0,0])"
            global PSE_A= pose_add (PSE_T, p[0,0,0.200,0,0,0])
          end
        end
      elif (4 == switch_2):
        $ 1538 "Case 4"
        $ 1539 "jig centrifuge racks"
        $ 1540 "define poses"
        $ 1541 "FRM_Reference≔ULM_Cent_Racks"
        global FRM_Reference=ULM_Cent_Racks
        $ 1542 "PSE_T≔get_pattern_pos_rectangle(JIG_Slot, 'X', [4,1], patternsize=[0.291,0])"
        global PSE_T=get_pattern_pos_rectangle(JIG_Slot, "X", [4,1], patternsize=[0.291,0])
        $ 1543 "If OBJ_Nbr≠0"
        if (OBJ_Nbr != 0):
          $ 1544 "PSE_T≔pose_trans(pose_trans(PSE_T, get_pattern_pos_rectangle(OBJ_Nbr, 'X', [3,3], patternsize=[0.060,0.060])),p[-0.030, -0.030,0,0,0,3.927])"
          global PSE_T= pose_trans ( pose_trans (PSE_T, get_pattern_pos_rectangle(OBJ_Nbr, "X", [3,3], patternsize=[0.060,0.060])),p[-0.030, -0.030,0,0,0,3.927])
        end
        $ 1545 "PSE_T≔pose_trans(PSE_T, GRP_Offset)"
        global PSE_T= pose_trans (PSE_T, GRP_Offset)
        $ 1546 "If Action≟1"
        if (Action == 1):
          $ 1547 "PSE_R≔pose_add(PSE_T, p[0,0,0.200,0,0,0])"
          global PSE_R= pose_add (PSE_T, p[0,0,0.200,0,0,0])
          $ 1548 "PSE_A≔pose_add(PSE_T, p[0,0,0.100,0,0,0])"
          global PSE_A= pose_add (PSE_T, p[0,0,0.100,0,0,0])
        else:
          $ 1549 "ElseIf Action≟2"
          if (Action == 2):
            $ 1550 "PSE_R≔pose_add(PSE_T, p[0,0,0.100,0,0,0])"
            global PSE_R= pose_add (PSE_T, p[0,0,0.100,0,0,0])
            $ 1551 "PSE_A≔pose_add(PSE_T, p[0,0,0.200,0,0,0])"
            global PSE_A= pose_add (PSE_T, p[0,0,0.200,0,0,0])
          end
        end
      elif (6 == switch_2):
        $ 1552 "Case 6"
        $ 1553 "Caps bin"
        $ 1554 "define poses"
        $ 1555 "'Drop cap'"
        # 'Drop cap'
        $ 1556 "FRM_Reference=ULM_Cap_Bin"
        FRM_Reference=ULM_Cap_Bin
        $ 1557 "PSE_T≔pose_RPY2RotVec(p[0,0,0,0,0,0])"
        global PSE_T=pose_RPY2RotVec(p[0,0,0,0,0,0])
        $ 1558 "PSE_T_H≔pose_add(PSE_T, p[0,0,-0.011,0,0,0])"
        global PSE_T_H= pose_add (PSE_T, p[0,0,-0.011,0,0,0])
        $ 1559 "PSE_A≔pose_trans(PSE_T, p[0,0,0.1,0,0,0])"
        global PSE_A= pose_trans (PSE_T, p[0,0,0.1,0,0,0])
        $ 1560 "PSE_R_H≔pose_add(PSE_T, p[0,0,0.100,0,0,0])"
        global PSE_R_H= pose_add (PSE_T, p[0,0,0.100,0,0,0])
        $ 1561 "PSE_R≔pose_add(PSE_T, p[0,0,0.100,0,0,0])"
        global PSE_R= pose_add (PSE_T, p[0,0,0.100,0,0,0])
      elif (7 == switch_2):
        $ 1562 "Case 7"
      elif (8 == switch_2):
        $ 1587 "Case 8"
        $ 1588 "NoK"
        $ 1589 "define poses"
        $ 1590 "'NoK'"
        # 'NoK'
        $ 1591 "FRM_Reference=ULM_NoK"
        FRM_Reference=ULM_NoK
        $ 1592 "PSE_T≔pose_RPY2RotVec(p[0,0,0,0,0,0])"
        global PSE_T=pose_RPY2RotVec(p[0,0,0,0,0,0])
        $ 1593 "PSE_A≔pose_trans(PSE_T, p[0,0,0.1,0,0,0])"
        global PSE_A= pose_trans (PSE_T, p[0,0,0.1,0,0,0])
        $ 1594 "PSE_R≔pose_add(PSE_T, p[0,0,0.100,0,0,0])"
        global PSE_R= pose_add (PSE_T, p[0,0,0.100,0,0,0])
      elif (9 == switch_2):
        $ 1595 "Case 9"
      elif (10 == switch_2):
        $ 1603 "Case 10"
      elif (11 == switch_2):
        $ 1611 "Case 11"
      elif (12 == switch_2):
        $ 1619 "Case 12"
      end
    elif (2 == switch_1):
      $ 1627 "Case 2"
      $ 1628 "Centrifuge"
      $ 1629 "'CHANGE THE REFERENCE TO THE FRAME TO MOVE IN'"
      # 'CHANGE THE REFERENCE TO THE FRAME TO MOVE IN'
      $ 1630 "define poses"
      $ 1631 "FRM_Reference≔FRM_Centrifuge"
      global FRM_Reference=FRM_Centrifuge
      $ 1632 "PSE_T≔GRP_Offset"
      global PSE_T=GRP_Offset
      $ 1633 "If Action≟8"
      if (Action == 8):
        $ 1634 "PSE_R≔pose_add(PSE_T, p[0,0,0.250,0,0,0])"
        global PSE_R= pose_add (PSE_T, p[0,0,0.250,0,0,0])
        $ 1635 "PSE_A≔pose_add(PSE_T, p[0,0,0.150,0,0,0])"
        global PSE_A= pose_add (PSE_T, p[0,0,0.150,0,0,0])
      else:
        $ 1636 "ElseIf Action≟7"
        if (Action == 7):
          $ 1637 "PSE_R≔pose_add(PSE_T, p[0,0,0.150,0,0,0])"
          global PSE_R= pose_add (PSE_T, p[0,0,0.150,0,0,0])
          $ 1638 "PSE_A≔pose_add(PSE_T, p[0,0,0.250,0,0,0])"
          global PSE_A= pose_add (PSE_T, p[0,0,0.250,0,0,0])
        end
      end
    elif (3 == switch_1):
      $ 1639 "Case 3"
      $ 1640 "Output"
      $ 1641 "'CHANGE THE REFERENCE TO THE FRAME TO MOVE IN'"
      # 'CHANGE THE REFERENCE TO THE FRAME TO MOVE IN'
      $ 1642 "define poses"
      $ 1643 "FRM_Reference≔Base_const"
      global FRM_Reference=p[0.0,0.0,0.0,0.0,0.0,0.0]
      $ 1644 "PSE_T≔p[0,0,0,0,0,0]"
      global PSE_T=p[0,0,0,0,0,0]
      $ 1645 "PSE_A≔pose_add(PSE_T, p[0,0,0.150,0,0,0])"
      global PSE_A= pose_add (PSE_T, p[0,0,0.150,0,0,0])
      $ 1646 "PSE_R≔pose_add(PSE_T, p[0,0,0.100,0,0,0])"
      global PSE_R= pose_add (PSE_T, p[0,0,0.100,0,0,0])
    elif (5 == switch_1):
      $ 1647 "Case 5"
      $ 1648 "Sarstedt Pickup Table"
      $ 1649 "'CHANGE THE REFERENCE TO THE FRAME TO MOVE IN'"
      # 'CHANGE THE REFERENCE TO THE FRAME TO MOVE IN'
      $ 1650 "Switch JIG"
      switch_2 = JIG
      $ 1651 "Case 7"
      if (7 == switch_2):
        $ 1664 "Sarstedt"
        $ 1665 "'CHANGE THE REFERENCE TO THE FRAME TO MOVE IN'"
        # 'CHANGE THE REFERENCE TO THE FRAME TO MOVE IN'
        $ 1671 "If TASK.ID≟10"
        if (TASK.ID == 10):
          $ 1672 "Frame & Position Params"
          $ 1673 "FRM_Reference = CAM_LM_SSRack"
          FRM_Reference = CAM_LM_SSRack
          $ 1674 "PSE_T≔uLM_SS_PickPlc"
          global PSE_T=uLM_SS_PickPlc
          $ 1675 "PSE_A≔pose_trans(PSE_T, p[0,0,0.1,0,0,0])"
          global PSE_A= pose_trans (PSE_T, p[0,0,0.1,0,0,0])
          $ 1676 "PSE_R≔pose_add(PSE_T, p[0,0,0.1,0,0,0])"
          global PSE_R= pose_add (PSE_T, p[0,0,0.1,0,0,0])
        end
      end
    elif (13 == switch_1):
      $ 1683 "Case 13"
      $ 1684 "Sarstedt Pickup Table"
      $ 1685 "'CHANGE THE REFERENCE TO THE FRAME TO MOVE IN'"
      # 'CHANGE THE REFERENCE TO THE FRAME TO MOVE IN'
      $ 1686 "Switch JIG"
      switch_2 = JIG
      $ 1687 "Case 7"
      if (7 == switch_2):
        $ 1700 "Bottle"
        $ 1701 "'CHANGE THE REFERENCE TO THE FRAME TO MOVE IN'"
        # 'CHANGE THE REFERENCE TO THE FRAME TO MOVE IN'
        $ 1707 "If TASK.ID≟43"
        if (TASK.ID == 43):
          $ 1708 "Frame & Position Params"
          $ 1710 "PSE_T≔uLM_SS_PickPlc"
          global PSE_T=uLM_SS_PickPlc
          $ 1711 "PSE_A≔pose_trans(PSE_T, p[0,0,0.1,0,0,0])"
          global PSE_A= pose_trans (PSE_T, p[0,0,0.1,0,0,0])
          $ 1712 "PSE_R≔pose_add(PSE_T, p[0,0,0.1,0,0,0])"
          global PSE_R= pose_add (PSE_T, p[0,0,0.1,0,0,0])
        end
      end
    end
    $ 1719 "Additional check"
    $ 1720 "If  not is_reachable(FRM_Reference,[PSE_A,PSE_A_H,PSE_T,PSE_T_H,PSE_R,PSE_R_H])"
    if (  not  is_reachable(FRM_Reference,[PSE_A,PSE_A_H,PSE_T,PSE_T_H,PSE_R,PSE_R_H])):
      $ 1721 "Error"
      $ 1722 "set_error(ERROR_POSE_NOT_REACHABLE)"
      set_error(ERROR_POSE_NOT_REACHABLE)
      $ 1723 "Action≔0"
      global Action=0
    end
    $ 1724 "'=========='"
    # '=========='
    $ 1725 "Switch Action"
    switch_1 = Action
    $ 1726 "Case 1"
    if (1 == switch_1):
      $ 1727 "Pick"
      $ 1728 "Action_Info≔'pick object'"
      global Action_Info="pick object"
      $ 1729 "do_transition(pose_trans(FRM_Reference, PSE_T), keep_rxry=OBJ_Picked)"
      do_transition( pose_trans (FRM_Reference, PSE_T), keep_rxry=OBJ_Picked)
      $ 1730 "EOAT"
      $ 1731 "If  not OBJ_Picked"
      if (  not  OBJ_Picked):
        $ 1732 "rq_move_and_wait_mm(GRP_Open_Pos)"
         rq_move_and_wait_mm (GRP_Open_Pos)
      end
      $ 1733 "If PSE_A_H≠PSE_Z"
      if (PSE_A_H != PSE_Z):
        $ 1734 "If JNT_Q≠JNT_Z"
        if (JNT_Q != JNT_Z):
          $ 1735 "movej(get_inverse_kin(pose_trans(FRM_Reference, PSE_A_H), qnear=JNT_Q), r=0.050)"
          movej(get_inverse_kin( pose_trans (FRM_Reference, PSE_A_H), qnear=JNT_Q), r=0.050)
        else:
          $ 1736 "Else" "noBreak"
          $ 1737 "movej(pose_trans(FRM_Reference, PSE_A_H), r=0.050)"
          movej( pose_trans (FRM_Reference, PSE_A_H), r=0.050)
        end
      end
      $ 1738 "If PSE_A≠PSE_Z"
      if (PSE_A != PSE_Z):
        $ 1739 "If JNT_Q≠JNT_Z"
        if (JNT_Q != JNT_Z):
          $ 1740 "movej(get_inverse_kin(pose_trans(FRM_Reference, PSE_A), qnear=JNT_Q), r=0.020)"
          movej(get_inverse_kin( pose_trans (FRM_Reference, PSE_A), qnear=JNT_Q), r=0.020)
        else:
          $ 1741 "Else" "noBreak"
          $ 1742 "movej(pose_trans(FRM_Reference, PSE_A), r=0.020)"
          movej( pose_trans (FRM_Reference, PSE_A), r=0.020)
        end
      end
      $ 1743 "MoveL"
      $ 1744 "If PSE_T_H≠PSE_Z"
      if (PSE_T_H != PSE_Z):
        $ 1745 "PSE_T_H" "breakAfter"
        movel(pose_trans(FRM_Reference, PSE_T_H), a=0.5, v=0.4, r=0.01)
      end
      $ 1746 "PSE_T" "breakAfter"
      movel(pose_trans(FRM_Reference, PSE_T), a=0.08, v=0.12)
      $ 1747 "EOAT"
      $ 1748 "rq_set_force_norm(50)"
       rq_set_force_norm (50)
      $ 1749 "rq_close_and_wait()"
       rq_close_and_wait ()
      $ 1750 "OBJ_Picked≔rq_is_object_detected()"
      global OBJ_Picked= rq_is_object_detected ()
      $ 1751 "If  not OBJ_Picked"
      if (  not  OBJ_Picked):
        $ 1752 "set_error(ERROR_NO_OBJECT_TO_PICK)"
        set_error(ERROR_NO_OBJECT_TO_PICK)
      end
      $ 1753 "EXTT"
      $ 1754 "Switch JIG"
      switch_2 = JIG
      $ 1755 "Case 1"
      if (1 == switch_2):
        $ 1756 "3FG"
        $ 1757 "If OBJ_Picked"
        if (OBJ_Picked):
          $ 1758 "Set GRP_3F_Open=On"
          set_standard_digital_out(5, True)
        end
      end
      $ 1759 "If PSE_R_H≠PSE_Z"
      if (PSE_R_H != PSE_Z):
        $ 1760 "PSE_R" "breakAfter"
        movel(pose_trans(FRM_Reference, PSE_R), a=0.5, v=0.4, r=0.01)
        $ 1761 "PSE_R_H" "breakAfter"
        movel(pose_trans(FRM_Reference, PSE_R_H), a=0.5, v=0.4)
      else:
        $ 1762 "Else" "noBreak"
        $ 1763 "PSE_R" "breakAfter"
        movel(pose_trans(FRM_Reference, PSE_R), a=0.5, v=0.4)
      end
    elif (2 == switch_1):
      $ 1764 "Case 2"
      $ 1765 "Place"
      $ 1766 "Action_Info≔'place object'"
      global Action_Info="place object"
      $ 1767 "do_transition(pose_trans(FRM_Reference, PSE_T), keep_rxry=OBJ_Picked)"
      do_transition( pose_trans (FRM_Reference, PSE_T), keep_rxry=OBJ_Picked)
      $ 1768 "EXTT"
      $ 1769 "Switch JIG"
      switch_2 = JIG
      $ 1770 "Case 1"
      if (1 == switch_2):
        $ 1771 "3FG"
        $ 1772 "If OBJ_Picked"
        if (OBJ_Picked):
          $ 1773 "Set GRP_3F_Open=On"
          set_standard_digital_out(5, True)
        end
      end
      $ 1774 "If PSE_A_H≠PSE_Z"
      if (PSE_A_H != PSE_Z):
        $ 1775 "If JNT_Q≠JNT_Z"
        if (JNT_Q != JNT_Z):
          $ 1776 "movej(get_inverse_kin(pose_trans(FRM_Reference, PSE_A_H), qnear=JNT_Q), r=0.050)"
          movej(get_inverse_kin( pose_trans (FRM_Reference, PSE_A_H), qnear=JNT_Q), r=0.050)
        else:
          $ 1777 "Else" "noBreak"
          $ 1778 "movej(pose_trans(FRM_Reference, PSE_A_H), r=0.050)"
          movej( pose_trans (FRM_Reference, PSE_A_H), r=0.050)
        end
      end
      $ 1779 "If PSE_A≠PSE_Z"
      if (PSE_A != PSE_Z):
        $ 1780 "If JNT_Q≠JNT_Z"
        if (JNT_Q != JNT_Z):
          $ 1781 "movej(get_inverse_kin(pose_trans(FRM_Reference, PSE_A), qnear=JNT_Q), r=0.020)"
          movej(get_inverse_kin( pose_trans (FRM_Reference, PSE_A), qnear=JNT_Q), r=0.020)
        else:
          $ 1782 "Else" "noBreak"
          $ 1783 "movej(pose_trans(FRM_Reference, PSE_A), r=0.020)"
          movej( pose_trans (FRM_Reference, PSE_A), r=0.020)
        end
      end
      $ 1784 "MoveL"
      $ 1785 "If PSE_T_H≠PSE_Z"
      if (PSE_T_H != PSE_Z):
        $ 1786 "PSE_T_H" "breakAfter"
        movel(pose_trans(FRM_Reference, PSE_T_H), a=0.5, v=0.4, r=0.01)
      end
      $ 1787 "PSE_T" "breakAfter"
      global move_thread_flag_1787=0
      thread move_thread_1787():
        enter_critical
        move_thread_flag_1787 = 1
        movel(pose_trans(FRM_Reference, PSE_T), a=0.05, v=0.09)
        move_thread_flag_1787 = 2
        exit_critical
      end
      move_thread_flag_1787 = 0
      move_thread_han_1787 = run move_thread_1787()
      while (True):
        local targetTcpDirection=get_target_tcp_speed()
        local stepsToRetract=tool_contact(direction=targetTcpDirection)
        if (stepsToRetract > 0):
          kill move_thread_han_1787
          stopl(0.5)
          $ 1788 "Until (tool_contact_detection)"
          break
        end
        sleep(1.0E-10)
        if (move_thread_flag_1787 > 1):
          join move_thread_han_1787
          break
        end
        sync()
      end
      $ 1789 "Force"
      sleep(0.02)
      zero_ftsensor()
      force_mode(FRM_Reference, [1, 1, 1, 0, 0, 0], [0.0, 0.0, 0.0, 0.0, 0.0, 0.0], 2, [0.1, 0.1, 0.01, 0.3490658503988659, 0.3490658503988659, 0.3490658503988659])
      $ 1790 "PSE_T" "noBreak"
      movel(pose_trans(FRM_Reference, PSE_T), a=0.04, v=0.07)
      end_force_mode()
      stopl(5.0)
      $ 1791 "EXTT"
      $ 1792 "Switch JIG"
      switch_2 = JIG
      $ 1793 "Case 1"
      if (1 == switch_2):
        $ 1794 "3FG"
        $ 1795 "If OBJ_Picked"
        if (OBJ_Picked):
          $ 1796 "Set GRP_3F_Open=Off"
          set_standard_digital_out(5, False)
          $ 1797 "Wait: 0.2"
          sleep(0.2)
        end
      end
      $ 1798 "EOAT"
      $ 1799 "rq_move_and_wait_mm(GRP_Open_Pos)"
       rq_move_and_wait_mm (GRP_Open_Pos)
      $ 1800 "OBJ_Picked≔rq_is_object_detected()"
      global OBJ_Picked= rq_is_object_detected ()
      $ 1801 "If PSE_R_H≠PSE_Z"
      if (PSE_R_H != PSE_Z):
        $ 1802 "PSE_R" "breakAfter"
        movel(pose_trans(FRM_Reference, PSE_R), a=0.5, v=0.4, r=0.01)
        $ 1803 "PSE_R_H" "breakAfter"
        movel(pose_trans(FRM_Reference, PSE_R_H), a=0.5, v=0.4)
      else:
        $ 1804 "Else" "noBreak"
        $ 1805 "PSE_R" "breakAfter"
        movel(pose_trans(FRM_Reference, PSE_R), a=0.5, v=0.4)
      end
    elif (3 == switch_1):
      $ 1806 "Case 3"
      $ 1807 "Push"
      $ 1808 "Action_Info≔'push'"
      global Action_Info="push"
    elif (4 == switch_1):
      $ 1809 "Case 4"
      $ 1810 "Pull"
      $ 1811 "Action_Info≔'pull'"
      global Action_Info="pull"
    elif (6 == switch_1):
      $ 1814 "Case 6"
      $ 1815 "Drop the cap"
      $ 1816 "If JNT_A≠[0,0,0,0,0,0]"
      if (JNT_A != [0,0,0,0,0,0]):
        $ 1817 "MoveJ"
        $ 1818 "JNT_A" "breakAfter"
        movej(JNT_A, a=1.3962634015954636, v=1.7453292519943295, r=0.02)
      else:
        $ 1819 "Else" "noBreak"
        $ 1820 "MoveJ"
        $ 1821 "PSE_A" "breakAfter"
        movej(pose_trans(FRM_Reference, PSE_A), a=1.3962634015954636, v=1.7453292519943295, r=0.02)
      end
      $ 1822 "MoveL"
      $ 1823 "PSE_T" "breakAfter"
      movel(pose_trans(FRM_Reference, PSE_T), a=0.05, v=0.09)
      $ 1824 "'ADD OPEN GRIPPER'"
      # 'ADD OPEN GRIPPER'
      # begin: URCap Program Node
      #   Source: Robotiq_Grippers, 3.17.0.105337, Robotiq Inc.
      #   Type: Gripper
      $ 1825 "Gripper Move10mm (1)"
      if not(gripper_connected[0]):
        popup("Gripper 1 must be connected to run this program.", "No connection", False, True, True)
      end
      if not(rq_is_gripper_activated("1")):
        popup("Gripper 1 is not activated. Go to Installation tab > Gripper to activate it and run the program again.", "Not activated", False, True, True)
      end
      rq_set_pos_spd_for(201, 0, 28, "1")
      rq_wait_pos_spe_for_request(201, 0, 28, "1")
      rq_go_to("1")
      rq_wait("1")
      # end: URCap Program Node
      $ 1826 "PSE_T_H" "breakAfter"
      movel(pose_trans(FRM_Reference, PSE_T_H), a=0.05, v=0.09)
      # begin: URCap Program Node
      #   Source: Robotiq_Grippers, 3.17.0.105337, Robotiq Inc.
      #   Type: Gripper
      $ 1827 "Gripper Move40mm (1)"
      if not(gripper_connected[0]):
        popup("Gripper 1 must be connected to run this program.", "No connection", False, True, True)
      end
      if not(rq_is_gripper_activated("1")):
        popup("Gripper 1 is not activated. Go to Installation tab > Gripper to activate it and run the program again.", "Not activated", False, True, True)
      end
      rq_set_pos_spd_for(63, 0, 28, "1")
      rq_wait_pos_spe_for_request(63, 0, 28, "1")
      rq_go_to("1")
      rq_wait("1")
      # end: URCap Program Node
      $ 1828 "PSE_R" "breakAfter"
      movel(pose_trans(FRM_Reference, PSE_R), a=0.5, v=0.4)
    elif (7 == switch_1):
      $ 1829 "Case 7"
      $ 1830 "Load"
      $ 1831 "Action_Info≔'load object'"
      global Action_Info="load object"
      $ 1832 "do_transition(pose_trans(FRM_Reference, PSE_T), keep_rxry=OBJ_Picked)"
      do_transition( pose_trans (FRM_Reference, PSE_T), keep_rxry=OBJ_Picked)
      $ 1833 "If PSE_A_H≠PSE_Z"
      if (PSE_A_H != PSE_Z):
        $ 1834 "If JNT_Q≠JNT_Z"
        if (JNT_Q != JNT_Z):
          $ 1835 "movej(get_inverse_kin(pose_trans(FRM_Reference, PSE_A_H), qnear=JNT_Q), r=0.050)"
          movej(get_inverse_kin( pose_trans (FRM_Reference, PSE_A_H), qnear=JNT_Q), r=0.050)
        else:
          $ 1836 "Else" "noBreak"
          $ 1837 "movej(pose_trans(FRM_Reference, PSE_A_H), r=0.050)"
          movej( pose_trans (FRM_Reference, PSE_A_H), r=0.050)
        end
      end
      $ 1838 "If PSE_A≠PSE_Z"
      if (PSE_A != PSE_Z):
        $ 1839 "If JNT_Q≠JNT_Z"
        if (JNT_Q != JNT_Z):
          $ 1840 "movej(get_inverse_kin(pose_trans(FRM_Reference, PSE_A), qnear=JNT_Q), r=0.020)"
          movej(get_inverse_kin( pose_trans (FRM_Reference, PSE_A), qnear=JNT_Q), r=0.020)
        else:
          $ 1841 "Else" "noBreak"
          $ 1842 "movej(pose_trans(FRM_Reference, PSE_A), r=0.020)"
          movej( pose_trans (FRM_Reference, PSE_A), r=0.020)
        end
      end
      $ 1843 "MoveL"
      $ 1844 "If PSE_T_H≠PSE_Z"
      if (PSE_T_H != PSE_Z):
        $ 1845 "PSE_T_H" "breakAfter"
        movel(pose_trans(FRM_Reference, PSE_T_H), a=0.5, v=0.4, r=0.01)
      end
      $ 1846 "PSE_T" "breakAfter"
      global move_thread_flag_1846=0
      thread move_thread_1846():
        enter_critical
        move_thread_flag_1846 = 1
        movel(pose_trans(FRM_Reference, PSE_T), a=0.05, v=0.09)
        move_thread_flag_1846 = 2
        exit_critical
      end
      move_thread_flag_1846 = 0
      move_thread_han_1846 = run move_thread_1846()
      while (True):
        local targetTcpDirection=get_target_tcp_speed()
        local stepsToRetract=tool_contact(direction=targetTcpDirection)
        if (stepsToRetract > 0):
          kill move_thread_han_1846
          stopl(0.5)
          $ 1847 "Until (tool_contact_detection)"
          break
        end
        sleep(1.0E-10)
        if (move_thread_flag_1846 > 1):
          join move_thread_han_1846
          break
        end
        sync()
      end
      $ 1848 "Force"
      sleep(0.02)
      zero_ftsensor()
      force_mode(FRM_Reference, [0, 1, 1, 0, 0, 1], [0.0, 0.0, 0.0, 0.0, 0.0, 0.0], 2, [0.1, 0.05, 0.02, 0.3490658503988659, 0.3490658503988659, 3.141592653589793])
      $ 1849 "PSE_T" "noBreak"
      movel(pose_trans(FRM_Reference, PSE_T), a=0.04, v=0.07)
      end_force_mode()
      stopl(5.0)
      $ 1850 "EOAT"
      $ 1851 "rq_move_and_wait_mm(GRP_Open_Pos)"
       rq_move_and_wait_mm (GRP_Open_Pos)
      $ 1852 "OBJ_Picked≔rq_is_object_detected()"
      global OBJ_Picked= rq_is_object_detected ()
      $ 1853 "If PSE_R_H≠PSE_Z"
      if (PSE_R_H != PSE_Z):
        $ 1854 "PSE_R" "breakAfter"
        movel(pose_trans(FRM_Reference, PSE_R), a=0.5, v=0.4, r=0.01)
        $ 1855 "PSE_R_H" "breakAfter"
        movel(pose_trans(FRM_Reference, PSE_R_H), a=0.5, v=0.4)
      else:
        $ 1856 "Else" "noBreak"
        $ 1857 "PSE_R" "breakAfter"
        movel(pose_trans(FRM_Reference, PSE_R), a=0.5, v=0.4)
      end
    elif (8 == switch_1):
      $ 1858 "Case 8"
      $ 1859 "Unload"
      $ 1860 "Action_Info≔'pick object'"
      global Action_Info="pick object"
      $ 1861 "do_transition(pose_trans(FRM_Reference, PSE_T), keep_rxry=OBJ_Picked)"
      do_transition( pose_trans (FRM_Reference, PSE_T), keep_rxry=OBJ_Picked)
      $ 1862 "EOAT"
      $ 1863 "If  not OBJ_Picked"
      if (  not  OBJ_Picked):
        $ 1864 "rq_move_and_wait_mm(GRP_Open_Pos)"
         rq_move_and_wait_mm (GRP_Open_Pos)
      end
      $ 1865 "If PSE_A_H≠PSE_Z"
      if (PSE_A_H != PSE_Z):
        $ 1866 "If JNT_Q≠JNT_Z"
        if (JNT_Q != JNT_Z):
          $ 1867 "movej(get_inverse_kin(pose_trans(FRM_Reference, PSE_A_H), qnear=JNT_Q), r=0.050)"
          movej(get_inverse_kin( pose_trans (FRM_Reference, PSE_A_H), qnear=JNT_Q), r=0.050)
        else:
          $ 1868 "Else" "noBreak"
          $ 1869 "movej(pose_trans(FRM_Reference, PSE_A_H), r=0.050)"
          movej( pose_trans (FRM_Reference, PSE_A_H), r=0.050)
        end
      end
      $ 1870 "If PSE_A≠PSE_Z"
      if (PSE_A != PSE_Z):
        $ 1871 "If JNT_Q≠JNT_Z"
        if (JNT_Q != JNT_Z):
          $ 1872 "movej(get_inverse_kin(pose_trans(FRM_Reference, PSE_A), qnear=JNT_Q), r=0.020)"
          movej(get_inverse_kin( pose_trans (FRM_Reference, PSE_A), qnear=JNT_Q), r=0.020)
        else:
          $ 1873 "Else" "noBreak"
          $ 1874 "movej(pose_trans(FRM_Reference, PSE_A), r=0.020)"
          movej( pose_trans (FRM_Reference, PSE_A), r=0.020)
        end
      end
      $ 1875 "MoveL"
      $ 1876 "If PSE_T_H≠PSE_Z"
      if (PSE_T_H != PSE_Z):
        $ 1877 "PSE_T_H" "breakAfter"
        movel(pose_trans(FRM_Reference, PSE_T_H), a=0.5, v=0.4, r=0.01)
      end
      $ 1878 "PSE_T" "breakAfter"
      movel(pose_trans(FRM_Reference, PSE_T), a=0.08, v=0.12)
      $ 1879 "Force"
      sleep(0.02)
      zero_ftsensor()
      force_mode(FRM_Reference, [1, 1, 0, 0, 0, 0], [0.0, 0.0, 0.0, 0.0, 0.0, 0.0], 2, [0.05, 0.05, 0.1, 0.3490658503988659, 0.3490658503988659, 0.3490658503988659])
      $ 1880 "EOAT" "noBreak"
      $ 1881 "rq_set_force_norm(50)" "noBreak"
       rq_set_force_norm (50)
      $ 1882 "rq_close_and_wait()" "noBreak"
       rq_close_and_wait ()
      $ 1883 "OBJ_Picked≔rq_is_object_detected()" "noBreak"
      global OBJ_Picked= rq_is_object_detected ()
      $ 1884 "If  not OBJ_Picked" "noBreak"
      if (  not  OBJ_Picked):
        $ 1885 "set_error(ERROR_NO_OBJECT_TO_PICK)" "noBreak"
        set_error(ERROR_NO_OBJECT_TO_PICK)
      end
      $ 1886 "If PSE_R_H≠PSE_Z" "noBreak"
      if (PSE_R_H != PSE_Z):
        $ 1887 "PSE_R" "noBreak"
        movel(pose_trans(FRM_Reference, PSE_R), a=0.5, v=0.4, r=0.01)
        $ 1888 "PSE_R_H" "noBreak"
        movel(pose_trans(FRM_Reference, PSE_R_H), a=0.5, v=0.4)
      else:
        $ 1889 "Else" "noBreak"
        $ 1890 "PSE_R" "noBreak"
        movel(pose_trans(FRM_Reference, PSE_R), a=0.5, v=0.4)
      end
      end_force_mode()
      stopl(5.0)
    elif (11 == switch_1):
      $ 1891 "Case 11"
    elif (12 == switch_1):
      $ 1928 "Case 12"
      $ 1929 "Decap"
      $ 1930 "Action_Info≔'decapping'"
      global Action_Info="decapping"
      $ 1931 "Set GRP_3F_Enable=On"
      set_standard_digital_out(4, True)
      $ 1932 "Set GRP_3F_Decap=On"
      set_standard_digital_out(3, True)
      $ 1933 "Force"
      sleep(0.02)
      zero_ftsensor()
      force_mode(tool_pose(), [0, 0, 1, 0, 0, 0], [0.0, 0.0, 5.0, 0.0, 0.0, 0.0], 2, [0.1, 0.1, 0.15, 0.3490658503988659, 0.3490658503988659, 0.3490658503988659])
      $ 1934 "check_decapping(offset=0.015, timeout=5, abort=CMD_Hold)" "noBreak"
      check_decapping(offset=0.015, timeout=5, abort=CMD_Hold)
      end_force_mode()
      stopl(5.0)
      $ 1935 "Set GRP_3F_Decap=Off"
      set_standard_digital_out(3, False)
      $ 1936 "Set GRP_3F_Enable=Off"
      set_standard_digital_out(4, False)
      $ 1937 "MoveL"
      $ 1938 "PSE_R" "breakAfter"
      movel(pose_trans(FRM_Reference, PSE_R), a=0.8, v=0.15)
    elif (13 == switch_1):
      $ 1939 "Case 13"
      $ 1940 "TMR_Barcode: Reset"
      TMR_Barcode = 0
      $ 1941 "Read"
      $ 1942 "TMR_Barcode: Start"
      TMR_Barcode_is_counting = True
      $ 1943 "If TMR_Barcode<PRM_TO_Read_BC"
      global thread_flag_1943=0
      thread Thread_if_1943():
        $ 1944 "KeyenceTrigger"
        $ 1945 "Set OClearResult=HI:Pulse 0.2"
        thread SinglePulse54():
          write_output_boolean_register(2, True)
          sleep(0.2)
          write_output_boolean_register(2, False)
        end
        singlePulse54 = run SinglePulse54()
        $ 1946 "Wait: 0.5"
        sleep(0.5)
        $ 1947 "Set OTriggerBarcode=Off"
        write_output_boolean_register(1, False)
        $ 1948 "Wait: 0.5"
        sleep(0.5)
        $ 1949 "Set OTriggerBarcode=On"
        write_output_boolean_register(1, True)
        $ 1950 "Wait: 0.5"
        sleep(0.5)
        $ 1951 "Preorient"
        $ 1952 "TMR_Barcode: Reset"
        TMR_Barcode = 0
        $ 1953 "If ICmdExctd"
        if (read_input_boolean_register(12)):
          $ 1954 "Set GRP_3F_Decap=On"
          set_standard_digital_out(3, True)
          $ 1955 "Set GRP_3F_Enable=On"
          set_standard_digital_out(4, True)
          $ 1956 "Loop ICmdExctd"
          while (read_input_boolean_register(12)):
            $ 1957 "KeyenceTrigger"
            $ 1958 "Set OClearResult=HI:Pulse 0.1"
            thread SinglePulse55():
              write_output_boolean_register(2, True)
              sleep(0.1)
              write_output_boolean_register(2, False)
            end
            singlePulse55 = run SinglePulse55()
            $ 1959 "Wait: 0.3"
            sleep(0.3)
            $ 1960 "Set OTriggerBarcode=Off"
            write_output_boolean_register(1, False)
            $ 1961 "Wait: 0.3"
            sleep(0.3)
            $ 1962 "Set OTriggerBarcode=On"
            write_output_boolean_register(1, True)
            $ 1963 "Wait: 0.1"
            sleep(0.1)
          end
        end
        $ 1964 "If  not ICmdExctd"
        if (  not  read_input_boolean_register(12)):
          $ 1965 "Set GRP_3F_Decap=On"
          set_standard_digital_out(3, True)
          $ 1966 "Set GRP_3F_Enable=On"
          set_standard_digital_out(4, True)
          $ 1967 "Wait ICmdExctd=HI"
          while (read_input_boolean_register(12) == False):
            sync()
          end
        end
        $ 1968 "Set GRP_3F_Decap=Off"
        set_standard_digital_out(3, False)
        $ 1969 "Set GRP_3F_Enable=Off"
        set_standard_digital_out(4, False)
        $ 1970 "OBJ_Brc_OK≔ True "
        global OBJ_Brc_OK=  True
        thread_flag_1943 = 1
      end
      if (TMR_Barcode<PRM_TO_Read_BC):
        global thread_handler_1943=run Thread_if_1943()
        while (thread_flag_1943 == 0):
          if not(TMR_Barcode<PRM_TO_Read_BC):
            kill thread_handler_1943
            thread_flag_1943 = 2
          else:
            sync()
          end
        end
      else:
        thread_flag_1943 = 2
      end
      if (thread_flag_1943 == 2):
        $ 1971 "Else" "noBreak"
        $ 1972 "exeption"
        $ 1973 "error"
        $ 1975 "OBJ_Brc_OK≔ False "
        global OBJ_Brc_OK=  False
      end
      $ 1976 "Set GRP_3F_Decap=Off"
      set_standard_digital_out(3, False)
      $ 1977 "Set GRP_3F_Enable=Off"
      set_standard_digital_out(4, False)
      $ 1978 "Set OTriggerBarcode=Off"
      write_output_boolean_register(1, False)
    elif (15 == switch_1):
      $ 1979 "Case 15"
      $ 1980 "Detect"
      $ 1981 "Action_Info≔'detect'"
      global Action_Info="detect"
    elif (30 == switch_1):
      $ 1982 "Case 30"
      $ 1983 "Shake"
      $ 1984 "Action_Info≔'shake'"
      global Action_Info="shake"
      $ 1985 "do_transition(pose_trans(FRM_Reference, PSE_T), keep_rxry=OBJ_Picked)"
      do_transition( pose_trans (FRM_Reference, PSE_T), keep_rxry=OBJ_Picked)
      $ 1986 "If PSE_A_H≠PSE_Z"
      if (PSE_A_H != PSE_Z):
        $ 1987 "If JNT_Q≠JNT_Z"
        if (JNT_Q != JNT_Z):
          $ 1988 "movej(get_inverse_kin(pose_trans(FRM_Reference, PSE_A_H), qnear=JNT_Q), r=0.050)"
          movej(get_inverse_kin( pose_trans (FRM_Reference, PSE_A_H), qnear=JNT_Q), r=0.050)
        else:
          $ 1989 "Else" "noBreak"
          $ 1990 "movej(pose_trans(FRM_Reference, PSE_A_H), r=0.050)"
          movej( pose_trans (FRM_Reference, PSE_A_H), r=0.050)
        end
      end
      $ 1991 "If PSE_A≠PSE_Z"
      if (PSE_A != PSE_Z):
        $ 1992 "If JNT_Q≠JNT_Z"
        if (JNT_Q != JNT_Z):
          $ 1993 "movej(get_inverse_kin(pose_trans(FRM_Reference, PSE_A), qnear=JNT_Q), r=0.020)"
          movej(get_inverse_kin( pose_trans (FRM_Reference, PSE_A), qnear=JNT_Q), r=0.020)
        else:
          $ 1994 "Else" "noBreak"
          $ 1995 "movej(pose_trans(FRM_Reference, PSE_A), r=0.020)"
          movej( pose_trans (FRM_Reference, PSE_A), r=0.020)
        end
      end
      $ 1996 "MoveL"
      $ 1997 "If PSE_T_H≠PSE_Z"
      if (PSE_T_H != PSE_Z):
        $ 1998 "PSE_T_H" "breakAfter"
        movel(pose_trans(FRM_Reference, PSE_T_H), a=0.5, v=0.4, r=0.01)
      end
      $ 1999 "PSE_T" "breakAfter"
      movel(pose_trans(FRM_Reference, PSE_T), a=0.08, v=0.12)
      $ 2000 "EXTT"
      $ 2001 "Comment"
      # Comment
      $ 2002 "MoveJ"
      $ 2003 "Waypoint_54" "breakAfter"
      movej(get_inverse_kin(Waypoint_54_p, qnear=Waypoint_54_q), a=1.3962634015954636, v=1.0471975511965976)
      $ 2004 "MoveJ"
      $ 2005 "Waypoint_77" "breakAfter"
      movej(get_inverse_kin(Waypoint_77_p, qnear=Waypoint_77_q), a=1.3962634015954636, v=1.0471975511965976)
      $ 2006 "MoveJ"
      $ 2007 "Waypoint_83" "breakAfter"
      movej(get_inverse_kin(Waypoint_83_p, qnear=Waypoint_83_q), a=1.3962634015954636, v=1.0471975511965976)
      $ 2008 "MoveJ"
      $ 2009 "Waypoint_84" "breakAfter"
      movej(get_inverse_kin(Waypoint_84_p, qnear=Waypoint_84_q), a=1.3962634015954636, v=1.0471975511965976)
      $ 2010 "If PSE_R_H≠PSE_Z"
      if (PSE_R_H != PSE_Z):
        $ 2011 "PSE_R" "breakAfter"
        movel(pose_trans(FRM_Reference, PSE_R), a=0.5, v=0.4, r=0.01)
        $ 2012 "PSE_R_H" "breakAfter"
        movel(pose_trans(FRM_Reference, PSE_R_H), a=0.5, v=0.4)
      else:
        $ 2013 "Else" "noBreak"
        $ 2014 "PSE_R" "breakAfter"
        movel(pose_trans(FRM_Reference, PSE_R), a=0.5, v=0.4)
      end
    elif (31 == switch_1):
      $ 2015 "Case 31"
      $ 2016 "Action_Info≔'Pick_Vial'"
      global Action_Info="Pick_Vial"
      $ 2017 "Pick_Vial"
      # begin: URCap Program Node
      #   Source: Robotiq_Grippers, 3.17.0.105337, Robotiq Inc.
      #   Type: Gripper
      $ 2018 "Gripper Open (1)"
      if not(gripper_connected[0]):
        popup("Gripper 1 must be connected to run this program.", "No connection", False, True, True)
      end
      if not(rq_is_gripper_activated("1")):
        popup("Gripper 1 is not activated. Go to Installation tab > Gripper to activate it and run the program again.", "Not activated", False, True, True)
      end
      rq_set_pos_spd_for(0, 82, 71, "1")
      rq_wait_pos_spe_for_request(0, 82, 71, "1")
      rq_go_to("1")
      rq_wait("1")
      # end: URCap Program Node
      $ 2019 "MoveJ"
      $ 2020 "Vial_above_1" "breakAfter"
      movej(get_inverse_kin(Vial_above_1_p, qnear=Vial_above_1_q), a=0.5235987755982988, v=0.4363323129985824, r=0.05)
      $ 2021 "MoveL"
      $ 2022 "Vial_pick_poi_1" "breakAfter"
      movel(Vial_pick_poi_1_p, a=0.5, v=0.1)
      # begin: URCap Program Node
      #   Source: Robotiq_Grippers, 3.17.0.105337, Robotiq Inc.
      #   Type: Gripper
      $ 2023 "Gripper Close (1)"
      if not(gripper_connected[0]):
        popup("Gripper 1 must be connected to run this program.", "No connection", False, True, True)
      end
      if not(rq_is_gripper_activated("1")):
        popup("Gripper 1 is not activated. Go to Installation tab > Gripper to activate it and run the program again.", "Not activated", False, True, True)
      end
      rq_set_pos_spd_for(255, 71, 84, "1")
      rq_wait_pos_spe_for_request(255, 71, 84, "1")
      rq_go_to("1")
      rq_wait("1")
      # end: URCap Program Node
      $ 2024 "MoveL"
      $ 2025 "Waypoint_86" "breakAfter"
      movel(Waypoint_86_p, a=0.5, v=0.1, r=0.05)
      $ 2026 "Home (Safe)"
      movej([-1.2302089344500047, -1.2969853503591224, -1.875639182904262, -1.539621866126728, 1.5731943360401213, -2.80099559440227], a=1.3962634015954636, v=1.0471975511965976)
    elif (32 == switch_1):
      $ 2027 "Case 32"
      $ 2029 "decap_Vial"
      $ 2030 "Set GRP_3F_Open=On"
      set_standard_digital_out(5, True)
      $ 2031 "MoveJ"
      $ 2032 "Waypoint_87" "breakAfter"
      movej(get_inverse_kin(Waypoint_87_p, qnear=Waypoint_87_q), a=0.5235987755982988, v=0.4363323129985824)
      $ 2033 "MoveL"
      $ 2034 "Vial_3FG_plac_1" "breakAfter"
      movel(Vial_3FG_plac_1_p, a=0.5, v=0.1)
      $ 2035 "Set GRP_3F_Open=Off"
      set_standard_digital_out(5, False)
      $ 2036 "Wait: 0.5"
      sleep(0.5)
      $ 2037 "MoveL"
      $ 2038 "Waypoint_88" "breakAfter"
      movel(Waypoint_88_p, a=0.5, v=0.1, r=0.05)
      $ 2039 "MoveJ"
      $ 2040 "cap_dump_1" "breakAfter"
      movej(get_inverse_kin(cap_dump_1_p, qnear=cap_dump_1_q), a=0.5235987755982988, v=0.4363323129985824)
      # begin: URCap Program Node
      #   Source: Robotiq_Grippers, 3.17.0.105337, Robotiq Inc.
      #   Type: Gripper
      $ 2041 "Gripper Open (1)"
      if not(gripper_connected[0]):
        popup("Gripper 1 must be connected to run this program.", "No connection", False, True, True)
      end
      if not(rq_is_gripper_activated("1")):
        popup("Gripper 1 is not activated. Go to Installation tab > Gripper to activate it and run the program again.", "Not activated", False, True, True)
      end
      rq_set_pos_spd_for(0, 255, 255, "1")
      rq_wait_pos_spe_for_request(0, 255, 255, "1")
      rq_go_to("1")
      rq_wait("1")
      # end: URCap Program Node
      $ 2042 "MoveJ"
      $ 2043 "Waypoint_89" "breakAfter"
      movej(get_inverse_kin(Waypoint_89_p, qnear=Waypoint_89_q), a=0.5235987755982988, v=0.4363323129985824, r=0.05)
      $ 2044 "MoveL"
      $ 2045 "Vial_3FG_plac_2" "breakAfter"
      movel(Vial_3FG_plac_2_p, a=0.5, v=0.1)
      # begin: URCap Program Node
      #   Source: Robotiq_Grippers, 3.17.0.105337, Robotiq Inc.
      #   Type: Gripper
      $ 2046 "Gripper Close (1)"
      if not(gripper_connected[0]):
        popup("Gripper 1 must be connected to run this program.", "No connection", False, True, True)
      end
      if not(rq_is_gripper_activated("1")):
        popup("Gripper 1 is not activated. Go to Installation tab > Gripper to activate it and run the program again.", "Not activated", False, True, True)
      end
      rq_set_pos_spd_for(255, 204, 255, "1")
      rq_wait_pos_spe_for_request(255, 204, 255, "1")
      rq_go_to("1")
      rq_wait("1")
      # end: URCap Program Node
      $ 2053 "Decap"
      $ 2054 "Action_Info≔'decapping'"
      global Action_Info="decapping"
      $ 2055 "Set GRP_3F_Enable=On"
      set_standard_digital_out(4, True)
      $ 2056 "Set GRP_3F_Decap=On"
      set_standard_digital_out(3, True)
      $ 2057 "Force"
      sleep(0.02)
      zero_ftsensor()
      force_mode(p[0.0,0.0,0.0,0.0,0.0,0.0], [0, 0, 1, 0, 0, 0], [0.0, 0.0, 1.0, 0.0, 0.0, 0.0], 2, [0.1, 0.1, 0.001, 0.3490658503988659, 0.3490658503988659, 0.3490658503988659])
      $ 2058 "check_decapping(offset=0.015, timeout=10, abort=CMD_Hold)" "noBreak"
      check_decapping(offset=0.015, timeout=10, abort=CMD_Hold)
      end_force_mode()
      stopl(5.0)
      $ 2059 "Set GRP_3F_Decap=Off"
      set_standard_digital_out(3, False)
      $ 2060 "Set GRP_3F_Enable=Off"
      set_standard_digital_out(4, False)
      $ 2061 "MoveL"
      $ 2062 "Waypoint_90" "breakAfter"
      movel(Waypoint_90_p, a=0.5, v=0.1, r=0.05)
      $ 2063 "MoveJ"
      $ 2064 "cap_dump_2" "breakAfter"
      movej(get_inverse_kin(cap_dump_2_p, qnear=cap_dump_2_q), a=0.5235987755982988, v=0.4363323129985824)
      # begin: URCap Program Node
      #   Source: Robotiq_Grippers, 3.17.0.105337, Robotiq Inc.
      #   Type: Gripper
      $ 2065 "Gripper Open (1)"
      if not(gripper_connected[0]):
        popup("Gripper 1 must be connected to run this program.", "No connection", False, True, True)
      end
      if not(rq_is_gripper_activated("1")):
        popup("Gripper 1 is not activated. Go to Installation tab > Gripper to activate it and run the program again.", "Not activated", False, True, True)
      end
      rq_set_pos_spd_for(0, 204, 255, "1")
      rq_wait_pos_spe_for_request(0, 204, 255, "1")
      rq_go_to("1")
      rq_wait("1")
      # end: URCap Program Node
      $ 2066 "MoveJ"
      $ 2067 "Waypoint_91" "breakAfter"
      movej(get_inverse_kin(Waypoint_91_p, qnear=Waypoint_91_q), a=0.5235987755982988, v=0.4363323129985824, r=0.036)
    elif (33 == switch_1):
      $ 2068 "Case 33"
      $ 2069 "Shake and liquid transfer"
      $ 2070 "MoveL"
      $ 2071 "Vial_liq_abov_1" "breakAfter"
      movel(Vial_liq_abov_1_p, a=0.5, v=0.1)
